(* IEC 61131-3 sources: SortJet_MasterSPS_Aufbau.fbsproj/06_Antriebe/Bosch Rexroth/Rexroth_ctrlX_Drive_Eckelmann_MC_V01_02_02.fb.st^, 26 files *)

(* ---- _Fehlerauswertung.act.st ---- *)
(* METADATA
{
	"v3Meta": {
		"objectGuid": "454009ed-4904-47be-a45e-86d01c03fc0f"
	}
}
*)
ACTION _Fehlerauswertung
/////////////////////////////////////////////////////////////////////////////////////////
/////////////////////////////////////////////////////////////////////////////////////////
// Fehlerauswertung
/////////////////////////////////////////////////////////////////////////////////////////
/////////////////////////////////////////////////////////////////////////////////////////
IF i_ui_Cia402_StatusWord.3 // Fehler am Umrichter aktiv
THEN
  Diagnose := DiagnoseAuswertung( wFehlernummer := udiErrorFromECat );
ELSE
  Diagnose := DiagnoseAuswertung( wFehlernummer := 0 );
END_IF

IF NOT i_ui_Cia402_StatusWord.3 AND NOT blInternerFehler AND blFehlerAktiv AND NOT blFreigabeEntziehenAktiv THEN
  Antriebsfehler.wlBausteinFehlerNr := cMotionFehler;
  blInternerFehler := TRUE;
END_IF

tonlFehlermeldungAusgeben(IN := ( blFehlerAktiv AND Diagnose.bError ) OR blInternerFehler , pt := T#1S);

rtl_Fehlermeldung(CLK := tonlFehlermeldungAusgeben.Q );

bpFehler := blFehlerAktiv AND ( Diagnose.bError (* OR Diagnose.bWarning *) OR blInternerFehler );

IF ( blInternerFehler ) THEN
  wlError := awlFehlerinformationen[4] := DWORD_TO_WORD(Antriebsfehler.wlBausteinFehlerNr);
ELSE
  awlFehlerinformationen[4] := DWORD_TO_WORD(Antriebsfehler.wlAntriebsFehler);
END_IF

IF ( rtl_Fehlermeldung.Q ) THEN

  awlFehlerinformationen[0] := stStationsNummern.NummerExtern;
  awlFehlerinformationen[1] := ppAntriebsInformationen.wpSchaltplanseite;
  awlFehlerinformationen[2] := ppAntriebsInformationen.wpSchaltplanReihe;
  awlFehlerinformationen[3] := ppAntriebsInformationen.wpSchaltschrank;

  IF ( blInternerFehler ) THEN
    SpsError( eFehler_Antrieb,
              wlError,
              stStationsNummern.NummerIntern,
              AutomatikkreisBestimmen(stStationsNummern.NummerSPS),
              awlFehlerinformationen );
  ELSE
    IF ( Diagnose.eType = eRexroth_Fehler_Error ) THEN
      SpsError( eFehler_Rexroth_Fehler + Diagnose.eErrorType,
                Diagnose.wFehlerNr,
                stStationsNummern.NummerIntern,
                AutomatikkreisBestimmen(stStationsNummern.NummerSPS),
                awlFehlerinformationen );
    // Wir loggen keine Warnungen
    // ELSIF ( Diagnose.eType = eRexroth_Fehler_Warning ) THEN
    //   SpsWarnung( eFehler_Rexroth_Warnung + Diagnose.eWarningType,
    //               Diagnose.wFehlerNr,
    //               stStationsNummern.NummerIntern,
    //               AutomatikkreisBestimmen(stStationsNummern.NummerSPS),
    //               awlErrorAdditional );
    END_IF
  END_IF

END_IF
END_ACTION

(* ---- _Statusword.act.st ---- *)
(* METADATA
{
	"v3Meta": {
		"objectGuid": "408b9d1a-1641-4edf-bb35-4e7a7361d31c"
	}
}
*)
ACTION _Statusword
/////////////////////////////////////////////////////////////////////////////////////////
/////////////////////////////////////////////////////////////////////////////////////////
// Aktuellen Status vom Antrieb auslesen
/////////////////////////////////////////////////////////////////////////////////////////
/////////////////////////////////////////////////////////////////////////////////////////
Status();

/////////////////////////////////////////////////////////////////////////////////////////
/////////////////////////////////////////////////////////////////////////////////////////
// Ist-Position auslesen
/////////////////////////////////////////////////////////////////////////////////////////
/////////////////////////////////////////////////////////////////////////////////////////
Istposition();

/////////////////////////////////////////////////////////////////////////////////////////
/////////////////////////////////////////////////////////////////////////////////////////
// Ist-Geschwindigkeit auslesen
/////////////////////////////////////////////////////////////////////////////////////////
/////////////////////////////////////////////////////////////////////////////////////////
IstGeschwindigkeit();

/////////////////////////////////////////////////////////////////////////////////////////
/////////////////////////////////////////////////////////////////////////////////////////
// Hardware Endschalter auslesen
/////////////////////////////////////////////////////////////////////////////////////////
/////////////////////////////////////////////////////////////////////////////////////////
// Rueckmeldung auch bei Quelle SPS aus dem Signal-Statuswort (im Umrichter parametriert)
IF ppAntriebsInformationen.stOptionen.eEndschalterQuelle <> Endschalterquelle_EN.KEINE THEN
  bpMaxSchalterBelegt := i_ui_Signal_StatusWord.1;
  bpMinSchalterBelegt := i_ui_Signal_StatusWord.0;
ELSE
  bpMinSchalterBelegt := FALSE;
  bpMaxSchalterBelegt := FALSE;
END_IF

/////////////////////////////////////////////////////////////////////////////////////////
/////////////////////////////////////////////////////////////////////////////////////////
// Erkennung ob und in welche Richtung der Antrieb verfährt
/////////////////////////////////////////////////////////////////////////////////////////
/////////////////////////////////////////////////////////////////////////////////////////
FahrrichtungErkennung();

/////////////////////////////////////////////////////////////////////////////////////////
/////////////////////////////////////////////////////////////////////////////////////////
// Status-Bits aus Antrieb / Motion holen
/////////////////////////////////////////////////////////////////////////////////////////
/////////////////////////////////////////////////////////////////////////////////////////
IF l_mc_ReadStatus.ErrorStop THEN
  l_mc_ReadAxisError( Axis := ppAntriebsInformationen.wAchsID , Enable := TRUE );
  blReadAxisErrorAktiv := TRUE;
ELSIF blReadAxisErrorAktiv THEN
  l_mc_ReadAxisError( Axis := ppAntriebsInformationen.wAchsID , Enable := FALSE );
  blReadAxisErrorAktiv := FALSE;
END_IF

blFehlerAktiv   := (  i_ui_Cia402_StatusWord.3 // Achsfehler
                     OR ( l_mc_ReadStatus.ErrorStop // MC Fehler
                          AND l_mc_ReadAxisError.Valid
                          AND NOT blFreigabeEntziehenAktiv ) // Aktiver Fehler aus MC_ReadAxisError
                     OR blInternerFehler ); // Fehler im Antriebsbaustein

bpIstReferenziert  := i_ui_Signal_StatusWord.3;
bpAchseSychron     := l_mc_GearIn.InGear (* AND l_mc_ReadStatus.SynchronizedMotion *);
bpBremseGeloest    := i_ui_Signal_StatusWord.15;

blSensoren[eSensoren.Sensor_1] := udipEingaengeUmrichter.cXG31_1_I_1;
blSensoren[eSensoren.Sensor_2] := udipEingaengeUmrichter.cXG31_2_I_2;
blSensoren[eSensoren.Sensor_3] := udipEingaengeUmrichter.cXG31_6_I_4;
blSensoren[eSensoren.Sensor_4] := udipEingaengeUmrichter.cXG31_7_I_5;
blSensoren[eSensoren.Sensor_5] := udipEingaengeUmrichter.cXG37_4_I_6;

// Sensorik vom Slave-gekoppelten Antrieb übernehmen - ggf kann man
IF IsBetweenWORD(wpSlaveNr, 0, 64) AND ( wpSlaveNr <> ppAntriebsInformationen.wAchsID ) THEN
  blSensoren[eSensoren.Sensor_6] := pgAntriebe[wpSlaveNr].udipEingaengeUmrichter.cXG31_1_I_1; // Slave Einlauf
  blSensoren[eSensoren.Sensor_7] := pgAntriebe[wpSlaveNr].udipEingaengeUmrichter.cXG31_2_I_2; // Slave Auslauf
  blSensoren[eSensoren.Sensor_8] := pgAntriebe[wpSlaveNr].udipEingaengeUmrichter.cXG31_6_I_4; // Slave Einlauf Vorab
  blSensoren[eSensoren.Sensor_9] := pgAntriebe[wpSlaveNr].udipEingaengeUmrichter.cXG31_7_I_5; // Slave Auslauf Vorab
ELSE
  blSensoren[eSensoren.Sensor_6] := FALSE;
  blSensoren[eSensoren.Sensor_7] := FALSE;
  blSensoren[eSensoren.Sensor_8] := FALSE;
  blSensoren[eSensoren.Sensor_9] := FALSE;
END_IF

bpMotionAktiv := ( NOT l_mc_ReadStatus.StandStill ) (* OR l_mc_ReadStatus.Disabled *);

bpAntrieblaeuft            := ( eBewegungsrichtung <> TE_Move_Direction.MD_STANDSTILL_E );
bpBewegungsrichtungPositiv := ( eBewegungsrichtung = TE_Move_Direction.MD_POSITIV_E );
bpBewegungsrichtungNegativ := ( eBewegungsrichtung = TE_Move_Direction.MD_NEGATIV_E );

bpKonstantfahrtAktiv       := l_mc_ReadStatus.ConstantVelocity;
bpBeschleunigungAktiv      := l_mc_ReadStatus.Accelerating;
bpVerzoegerungAktiv        := l_mc_ReadStatus.Decelerating;

bpReglerBereit      := ( PowerSupplyStatus.15 AND PowerSupplyStatus.14 AND PowerSupplyStatus.6 AND PowerSupplyStatus.4 )
                       OR ( i_ui_Cia402_StatusWord.0 AND i_ui_Cia402_StatusWord.1 AND i_ui_Cia402_StatusWord.2 );

// Min- und Max-Position bestimmen
rlSoftwareLimitMin := TO_REAL(l_ts_MKAxisConfig.lrSoftwareLimitNegative);
rlSoftwareLimitMax := TO_REAL(l_ts_MKAxisConfig.lrSoftwareLimitPositive);
rpMinPosition := rlSoftwareLimitMin;
rpMaxPosition := rlSoftwareLimitMax;

// Externe Software-Endschalter koennen die MK-Grenzen nur weiter eingrenzen
// 0 bedeutet: kein zusaetzlicher externer Endschalter aktiv

// Min nur enger setzen, nie erweitern
IF rpMinSwEsEingrenzung <> 0 THEN
  IF ( rlSoftwareLimitMin = 0 ) OR ( rpMinSwEsEingrenzung >= rlSoftwareLimitMin ) THEN
    rpMinPosition := rpMinSwEsEingrenzung;
  END_IF
END_IF

// Max nur enger setzen, nie erweitern
IF rpMaxSwEsEingrenzung <> 0 THEN
  IF ( rlSoftwareLimitMax = 0 ) OR ( rpMaxSwEsEingrenzung <= rlSoftwareLimitMax ) THEN
    rpMaxPosition := rpMaxSwEsEingrenzung;
  END_IF
END_IF

// Widerspruch im Ergebnis (Min > Max):
// externe Eingrenzung komplett verwerfen und MK-Grenzen beibehalten
IF rpMinPosition > rpMaxPosition THEN
  rpMinPosition := rlSoftwareLimitMin;
  rpMaxPosition := rlSoftwareLimitMax;
END_IF

blSoftwareLimitAktiv := ( rpMinPosition <> 0 ) OR ( rpMaxPosition <> 0 );

bpAntriebFreigegeben := (     l_mc_Power.Enable
                          AND l_mc_Power.Status );

rpPositionMesstaster1Positiv := TO_REAL(TO_LREAL(diTouchProbe1Pos) / l_ts_MKAxisConfig.lrIncrementsPerDistance * l_ts_MKAxisConfig.lrDistance);
rpPositionMesstaster1Negativ := TO_REAL(TO_LREAL(diTouchProbe1Neg) / l_ts_MKAxisConfig.lrIncrementsPerDistance * l_ts_MKAxisConfig.lrDistance);
rpPositionMesstaster2Positiv := TO_REAL(TO_LREAL(diTouchProbe2Pos) / l_ts_MKAxisConfig.lrIncrementsPerDistance * l_ts_MKAxisConfig.lrDistance);
rpPositionMesstaster2Negativ := TO_REAL(TO_LREAL(diTouchProbe2Neg) / l_ts_MKAxisConfig.lrIncrementsPerDistance * l_ts_MKAxisConfig.lrDistance);

bpHaupschalter400VEin := ppAntriebsInformationen.stOptionen.bVersorgungUeberXVR OR PowerSupplyStatus.4;

/////////////////////////////////////////////////////////////////////////////////////////
/////////////////////////////////////////////////////////////////////////////////////////
// Eingaenge vom Umrichter auslesen
/////////////////////////////////////////////////////////////////////////////////////////
/////////////////////////////////////////////////////////////////////////////////////////
bpLS_150F02_230V := ppAntriebsInformationen.stOptionen.bVersorgungUeberXVR OR udipEingaengeUmrichter.cXG31_3_I_3; // Eingang Leitungsschutzschalter 230V OK

// Ausgangssignale in diesem Normalzyklus uebernehmen, ins Steuerwort schreibt _Steuerwort
wlAusgaengeUmrichter := wpAusgaengeUmrichter;
END_ACTION

(* ---- _Steuerwort.act.st ---- *)
(* METADATA
{
	"v3Meta": {
		"objectGuid": "2cb5236d-2c9d-4e67-a004-d0a59f43b200"
	}
}
*)
ACTION _Steuerwort
// Alle Steuerwort-Bits werden ausschliesslich in dieser Aktion beschrieben.

// Externe Endschalter nur bei Quelle SPS weitergeben, sonst Frei-Pegel (Oeffner: TRUE = frei)
blEndschalterAusSPS := FALSE;
IF __ISVALIDREF(ppAntriebsInformationen) THEN
  blEndschalterAusSPS := ppAntriebsInformationen.stOptionen.eEndschalterQuelle = Endschalterquelle_EN.SPS;
END_IF

SignalSteuerWort.0  := blReferenzLoeschen;
SignalSteuerWort.1  := wlAusgaengeUmrichter.3;
SignalSteuerWort.2  := wlAusgaengeUmrichter.4;
SignalSteuerWort.3  := wlAusgaengeUmrichter.5;
SignalSteuerWort.4  := wlAusgaengeUmrichter.6;
SignalSteuerWort.5  := wlAusgaengeUmrichter.7;
SignalSteuerWort.6  := wlAusgaengeUmrichter.8;
SignalSteuerWort.7  := wlAusgaengeUmrichter.9;
SignalSteuerWort.8  := wlAusgaengeUmrichter.10;
SignalSteuerWort.9  := NOT blEndschalterAusSPS OR bpEndschalterMaxExtern;
SignalSteuerWort.10 := NOT blEndschalterAusSPS OR bpEndschalterMinExtern;
SignalSteuerWort.11 := FALSE;
SignalSteuerWort.12 := FALSE;
SignalSteuerWort.13 := FALSE;
SignalSteuerWort.14 := blReferenzSetzen;
SignalSteuerWort.15 := blBremseLoesen;
END_ACTION

(* ---- A_Changelog.act.st ---- *)
(* METADATA
{
	"v3Meta": {
		"objectGuid": "3ad406ab-889e-4d0d-be2f-76f9c9ecfe4e"
	}
}
*)
{attribute 'excludefrombuild'}
ACTION A_Changelog
(* !!! VERSIONSÄNDERUNGEN WERDEN HIER DETAILLIERT DOKUMENTIERT !!!

- 2025-07-02 - V01_00_00:
  - Entwicklung des Bausteins; Erste Version die Freigegeben wird/wurde

- 2025-10-10 - V01_00_01: Marc Wiegran
  - Änderung des Baustein. Damit die Visualisierung Antriebe_Verfahren weiterhin genutzt werden kann muss in den Schrittketten auf l_mc_power.Enable und nicht auf bpFreigabe geschaut werden.
    l_mc_power.Enable wird aus bpFreigabe und bpFrigabeErzingen, sodass wir nicht mehr in einen Internen Fehler laufen
  - Änderung des Bausteins Damit auch auf die gemeldeten zustände der Hardwarefreigabe geschaut wird wurde in den Schrittketten das l_mc_power.Status durch Regler bereit ersetzt

- 2025-10-15 - V01_00_02: Tobias Brekerbohm
  - Korrektur Vergleich der Software Endschalter - wenn beide 0 dann ansehen als wären keine Aktiv
  - Korrektur bpReglerBereit - Bei Achsen im Zwischenkreis kommen die Bits nicht entsprechend anderer Achsen
    Hier muss auf das CiA Status Word geschaut werden. Zu Prüfen ist, ob das bei den normalen Achsen auch ggf. schon ausreicht
  - Anpassungen / Korrekturen Rotative Achsen

- 2025-10-16 - V01_00_03: Tobias Brekerbohm
  - Korrektur dauernde Neuberechnung der Zielposition bei relativer Positionierung

- 2025-10-17 - V01_00_04: Marc Wiegran
  - Korrektur der Eingangsbits der Langsamfahrnocken auch CoE

- 2025-10-21 - V01_00_05: Marc Wiegran
  - Bei Geschwindigkeitsänderung bei der Messfahrt wird in Step 325 gesprungen um die MC_MOVE_Velocity neu zu starten und nicht wie vorher in 300, da dort erneut die Startbedingungen gepürft werden

- 2025-10-21 - V01_00_06: Marc Wiegran
  - Warteschritt 250 hinzugefgt um sicherzustellen, das die Softwarefreigabe vor Bewegungsstart erteilt wurde noch zu testen ob es die Fehler 6 der MC-Bausteine behebt
  - Schreiben der MC_Home-Fehler-ID in die dafür vorgesehene Variable

- 2025-10-22 - V01_00_07: Marc Wiegran
  - Entfernen des Warteschritt 250, statt dessen wird im Schritt 100 auf l_mc_Power.Status geschaut und Timerüberwacht wird dort ein Fehler ausgeworfen.
      - Enable := Freigabe setzten; Status := Freigabe wurde erfolgreich gesetzt
  - Entfernen der Überprüfung der aktuellen antriebsposition <100 nach der Referenz
      - die Querfahrten haben einen absoluten Referenzoffset von >100, sodass dies andernfalls nicht klappt

- 2025-10-28 - V01_00_08: Tobias Brekerbohm
  - State-Machine achtet nun auf NOT Valid als aller erstes
  - Vergessener Warteschritt 250 aus 1.00.06 der bei der Entfernung in 1.00.07 vergessen wurde zusätzlich entfernt

- 2025-11-11 - V01_00_09: Tobias Brekerbohm
  - Fehlerhaftes ABS setzen von Messergebnissen bei Scheibenmessungen entfernt

- 2025-11-13 - V01_00_10: Tobias Brekerbohm
  - Reset von Ref-Bezug löschen Bit hat gefehlt

- 2025-11-24 - V01_00_11: Tobias Brekerbohm
  - Fehlender Reset von Softwarefreigabe-Timer korigiert
  - An vielen Stellen wurde immernoch auf l_mc_Power.Enable geschaut für den Fehler der Softwarefreigabe statt auf l_mc_Power.Status

- 2026-12-10 - V01_00_12: Tobias Brekerbohm
  - Bei festen Zielpositionen werden keine mm/grad mehr aufaddiert, es werden hart die Grenzwerte aus dem EConSET genommen und nicht mehr schöngerechnet
  - Bei einer Zielpos außerhalb der Grenzen wird nun ein Fehler geworfen, statt die Zielpos stillschweigend zu begrenzen
  - Statt dauernd auf die MK Variablen zu schauen, welche noch konvertiert werden muss, wird nun direkt auf die rpMin- und rpMaxPosition geschaut

- 2026-12-10 - V01_00_13: Tobias Brekerbohm
  - bpAchseSychron schaut nicht länger auf l_mc_ReadStatus.SynchronizedMotion da das Signal aus dem Status gelegentlich geflackert hat

- 2026-12-10 - V01_00_14: Tobias Brekerbohm
  - ReadAxisError wurde nicht aufgerufen
  - Fehlerauswertung bei Fehler aus dem MotionKernel (F 108) bei kein Fehler vom Regler und kein internen Fehler

- 2026-03-12 - V01_00_15: Tobias Brekerbohm
  - Berechnung Ruckzeit bei Langsamfahrt fehlerhaft

- 2026-03-17 - V01_00_16: Tobias Brekerbohm
  - Handplus / Handminus / Restweg-Suchfahrt beachten nun die Software-Endschalter und bremsen vor Erreichen anhand der aktuellen Bremsposition ab
  - Ein Neustart in Richtung eines bereits ueberschrittenen Software-Endschalters wird unterbunden

- 2026-03-19 - V01_00_17: Tobias Brekerbohm
  - Neue Eingaben rpMinSwEsEingrenzung/rpMaxSwEsEingrenzung ergaenzen eine externe Eingrenzung der Software-Endschalter
  - Externe Limits duerfen den MK-Bereich nur enger machen und nicht erweitern
  - Alle Bewegungsarten pruefen neue Zielpositionen und Bremsgrenzen gegen die aktiven Min-/Max-Grenzen

- 2026-03-22 - V01_00_18: Tobias Brekerbohm
  - Antriebssimulation für SPS Simulation (ungetestet)

- 2026-03-24 - V01_00_19: Tobias Brekerbohm
  - XG37-1 und XG37-2 (eigentlich als Eingänge genutzt) optional auch als Ausgänge nutzbar (Benötigt Parameteränderung am Antrieb!!!)

- 2026-03-27 - V01_00_20: Tobias Brekerbohm
  - Neuer Eingang bpFreigabeEntziehenAnhalten fuer kontrollierten Freigabeentzug mit Halt ohne Schrittketten-Reset
  - Bei aktivem Freigabeentzug wird die Achse angehalten, danach die Power entzogen und nach Signalrueckkehr automatisch ohne externen Trigger fortgesetzt
  - Motion-Fehlerauswertung unterdrueckt erwartete ErrorStop-Meldungen waehrend aktivem Freigabeentzug
  - Beim Wiederanlauf nach Freigabeentzug werden laufende Schrittketten auf Execute-Startschritte remappt, damit Bewegungen sicher neu starten
  - Kein ungewollter Schrittketten-Reset bei Signalrueckkehr waehrend aktivem MC_Stop (rtlStop-Kante abgesichert)

- 2026-06-12 - V01_01_00: Tobias Brekerbohm
  - Globaler Override für die Achsgeschwindigkeit - Prozentual zu ändern. Neuer Input rpOverride 0-100
  - Taktzeitoptimierung: Flankenerkennung der Sensoren direkt im Antriebsbaustein ohne zusaetzlichen FB-Aufruf
  - Taktzeitoptimierung: Stillstandsposition nur bei aktiver Software-Endschalter-Bremswegueberwachung berechnen
  - Taktzeitoptimierung: MC_ReadAxisError nur im ErrorStop und einmalig zum Deaktivieren aufrufen
  - S277 Bit 12 wird geprüft, mit Fehlermeldung wenn nicht = 1
  - Bei aktivierter Langsamfahrtnocke wird nicht auf Langsame Geschwindigkeit gestellt, wenn die Achse beim belegen der Nocke/Laser gerade am Verzögern ist.
     Würden wir während der Verzögerung die Geschwindigkeit reduzieren, würde der Verfahrbefehl abgebrochen und neu geschrieben werden in den MotionKernel.
     Dabei verlieren wir Zeit und die Achse würde ihre Zielposition überfahren.
  - Restweg positionierung kann nun auch auf Achsen Restweg fahren, die per wpSlave angegeben werden. Z. b. Greifer auf Riemen-Sensorik (Sensor 6-9)
  - Gravierender Fehler bei der Langsamfahrt behoben: Shuttle überfährt seine Position massiv bei aktiver Langsamfahrt weil die Ruckzeit umgerechnet wurde und dadurch
    die Zielposition nicht mehr erreicht werden kann und somit überschwingt
  - Fehler behoben, dass blInternerFehler erst nach einem 2. Reset zurückgesetzt wurde. MotionFehler brauchten dadurch immer 2 Resets

- 2026-07-07 - V01_01_01: Tobias Brekerbohm
  - Fehler bei Zuweisung von Beschleunigung und Verzögerung behoben.

- 2026-08-04 - V01_01_02: Tobias Brekerbohm
  - Restwegmessung während der Absolutfahrt ermöglicht und Messung mehrerer aufeinanderfolgender Scheiben korrigiert.
  - Messergebnis der Restwegmessung wird immer positiv ausgegeben.

- 2026-08-05 - V01_01_03: Marc Wiegran und Tobias Brekerbohm
  - Korrektur zuweisung rpMessergbnis - Messergebnis war erst einen Zyklus nach erfolgreicher Messung im Statusword
  - Messergebnis der Längenmessung wird wieder negativ ausgegeben, da der Scheibenmessung_FB darauf ausgelegt ist den so zu erhalten

- 2026-09-25 - V01_01_04: Tobias Brekerbohm
  - Langsamfahrt begrenzt die Geschwindigkeit ueber MC_SetOverride auf 10 % der konfigurierten Maximalgeschwindigkeit.
  - Der externe rpOverride bleibt wirksam; Bewegungsbefehle werden fuer Langsamfahrt nicht mehr neu geschrieben.
  - Bei kurz erkanntem Stillstand bleibt aktive Langsamfahrt erhalten, solange eine Langsamfahrtnocke belegt ist.
  - Langsamfahrt-Bedingung in Nockenerkennung, Aktivierung und Halten aufgeteilt; Verhalten unveraendert.

- 2026-10-14 - V01_01_05: Tobias Brekerbohm:
  - FreigabeEntziehen_Wiederanlauf: MC_Stop wird auch ausgeloest, wenn der Antrieb laut MC-Status nicht im Stillstand ist (bisher nur ueber bpAntrieblaeuft -> bei Anlauf/langsamer Fahrt kein Stop und evtl. Power-Entzug waehrend der Fahrt)
  - FreigabeEntziehen_Wiederanlauf: tonlSoftwareFreigabe/tonlHardwareFreigabe werden waehrend des Halts zurueckgesetzt (Haltezeit zaehlt nicht als Timeout der eingefrorenen Schrittkette)

- 2026-10-17 - V01_02_00: Tobias Brekerbohm, Claude
  - Ruck (Jerk) für lineare und rotative Achsen überarbeitet: Kurze Fahrten nutzen von Anfang an den kleineren Jerk. Lange Fahrten starten mit dem Beschleunigungs-Jerk und wechseln bei erreichter Fahrgeschwindigkeit auf den Brems-Jerk. Der Brems-Jerk kann größer oder kleiner sein.
  - Ob eine Fahrt kurz oder lang ist, wird aus Strecke, Geschwindigkeit, Beschleunigung, Verzögerung und Ruckzeit berechnet. Die Ruckzeitbegrenzung aus EConSet wird berücksichtigt.
  - Der Wechsel auf den Brems-Jerk erfolgt nur einmal pro Fahrt. Parameteränderungen und eine Freigabepause schalten nicht wieder in die Beschleunigungsphase zurück.
  - Stoppen verwendet grundsätzlich den Brems-Jerk. Beim Abbruch während der Beschleunigung wird mindestens der Beschleunigungs-Jerk und der Jerk des laufenden Fahrbefehls verwendet. Dieser bleibt bis zum Ende des Stops erhalten, auch wenn die Schrittkette zurückgesetzt wird.
  - Die Jerk-Auswahl wird gemeinsam für Absolut-, Relativ-, Hand-, Mess-, Restweg- und Synchronfahrten verwendet. Strecken werden passend zum Achstyp in Millimetern oder Grad berechnet.

- 2026-10-19 - V01_02_01: Claude
  - Simulation (bgSPS_SIMULATION): MK-Konfiguration wird jetzt auch im Simulationsmodus geladen (MK_GetAxisConfiguration). Vorher blieb l_ts_MKAxisConfig leer und die Achsen liefen mit den Notfall-Grenzen +-1000.
  - Simulation: rlGeschwindigkeit/rlBeschleunigung/rlVerzoegerung werden jetzt wie in Pruefe_Inputs_Langsamfahrt aus den Eingaengen gebildet und auf die MK-Maximalwerte begrenzt. Vorher waren sie im Simulationsmodus immer 0, die Achsen fuhren daher immer mit den Fallback-Werten (200 / 800).
  - Simulation: rpOverride wirkt jetzt auch auf die simulierte Geschwindigkeit.
  - Simulation: Scheibenmessung (SCHEIBENMESSUNG) und Restwegmessung liefern jetzt ein Messergebnis. Mangels Glasmodell gilt eine virtuelle Scheibenlaenge (globale Variable rgSimScheibenlaenge, Standard 1000 mm):
    Die Messung ist abgeschlossen, wenn die Achse seit Messstart (bzw. seit der ersten Flanke bei Restweg) diese Strecke verfahren hat. Vorzeichen wie im Echtbetrieb angenommen: Scheibenmessung negativ (positiv bei bpDrehrichtungsumkehrMessung), Restweg positiv.
    Die Messfahrt laeuft wie im Echtbetrieb immer in positive Richtung. bpMessungOk/bpMessungFehlerhaft/rpMessErgebnis bleiben bis zum Betriebsartenwechsel gespeichert (vorher nur 1 Zyklus).
  - Simulation: Neuer Eingang rpSimMessErgebnis (nur Simulation): Station gibt das Ergebnis der Scheibenmessung vor. Echtbetrieb-Konvention (aus Scheibenmessung_FB): Ergebnis = Scheibenlaenge - Messstrecke, Glaslaenge = ABS(Messstrecke + Ergebnis).
    Die Messfahrt dauert so lange wie der Betrag des Ergebnisses. Ist der Eingang 0, gilt weiter die virtuelle Scheibenlaenge rgSimScheibenlaenge (Vorzeichen negativ).
  - Simulation: bpBremseLoesen setzt SignalSteuerWort.15 (nur mit bpBremseLoesenFreigabe, sonst Fehler) und meldet bpBremseGeloest nach 300 ms zurueck.
  - Simulation: bpAbsolutSetzen durchlaeuft wie im Echtbetrieb Referenz loeschen -> setzen -> bpAbsolutSetzenDone.
  - Simulation: Langsamfahrnocken (bpAktiviereLangsamfahrtNocke) sind jetzt Low-aktiv (FALSE = belegt) wie im Echtbetrieb, an den Wegenden positioniert; bpLangsamfahrenAktiv begrenzt die Geschwindigkeit auf 10 % der MK-Maximalgeschwindigkeit.
  - Simulation: Abbildung Sensor -> Umrichter-Eingang wie im Echtbetrieb (Sensor_3 = XG31_6, Sensor_4 = XG31_7, Sensor_5 = XG37_4; vorher um eine Stelle verschoben). Sensor_6..9 kommen wie im Echtbetrieb vom Slave-Antrieb (wpSlaveNr).

- 2026-10-31 - V01_02_02: Tobias Brekerbohm, Claude
  Hinweis: Die Nummer V01_01_05 wurde in zwei parallelen Zweigen doppelt vergeben: 2026-10-14 TB (FreigabeEntziehen_Wiederanlauf) und 2026-10-06 Daniel Vogelsang.
  Dieser Stand baut auf V01_02_01 auf und uebernimmt die Punkte aus dem zweiten Zweig (V01_01_05 vom 2026-10-06). Ruck-Profil, StopVerwaltung und Simulation bleiben wie in V01_02_01.
  - Steuerwort-Bits zentral in _Steuerwort zusammengefasst; Referenz- und Bremsenbefehle ueber interne BOOL-Merker. _Steuerwort laeuft auch vor den RETURN-Pfaden (ausser Achse 65).
  - Neue Struktur stOptionen (Antrieb_Optionen_ST) in AntriebsInformationen; ersetzt bpHardwareLimits und bpBremseLoesenFreigabe.
  - Endschalterquelle (eEndschalterQuelle): KEINE, UMRICHTER (Signal-Statuswort Bit 0 = Min, Bit 1 = Max) oder SPS.
  - Quelle SPS: Neue Eingaenge bpEndschalterMinExtern/bpEndschalterMaxExtern auf Signal-Steuerwort Bit 10 (Min) und Bit 9 (Max). Oeffner, TRUE = frei, Default TRUE fuer eine nicht vorhandene Seite.
    Bei anderer Quelle bleiben Bit 9/10 auf TRUE. bpMinSchalterBelegt/bpMaxSchalterBelegt kommen auch bei Quelle SPS aus dem Signal-Statuswort.
    Korrektur zum zweiten Zweig: Dort stehen Min/Max in Deklaration und Changelog vertauscht, gesendet wird Bit 9 = Max, Bit 10 = Min.
  - XVR-Modus (bVersorgungUeberXVR): brueckt bpHaupschalter400VEin und bpLS_150F02_230V, ersetzt die festen OR TRUE aus dem zweiten Zweig.
  - BETRIEBSART_MasterSlave Schritt 1000: bpDone wurde per Vergleich gebildet und war dadurch TRUE, obwohl die Achse nicht synchron war bzw. ein Fehler anstand. Jetzt bpDone := l_mc_GearIn.InGear, in den Fehlerzweigen bpDone := FALSE.
  - Defaults setzt bpDone := FALSE. Vorher blieb ein altes bpDone waehrend Busausfall stehen und ein Reset-Auftrag galt sofort als fertig.
  - tonlMaxZeitStatusUngueltig wird jeden Zyklus vor der State Machine aufgerufen und in Defaults zurueckgesetzt. Vorher wurde er nie zurueckgesetzt und eine spaetere kurze Statusstoerung loeste sofort einen Stop aus.
  - BETRIEBSART_Reset Schritt 250: l_mc_Reset.Error wird bewusst nicht ausgewertet. Der Changelog des zweiten Zweigs nennt diesen Punkt, der Code ist dort aber zu Recht auskommentiert.
  - BETRIEBSART_Reset: Neuer Schritt 260, wartet nach MC_Reset 1 s, bevor bei weiter anstehendem Fehler der Reset per CoE laeuft (aus dem zweiten Zweig).
  - _Statusword und Simulation: Widerspruchspruefung der Software-Endschalter auf das Ergebnis (rpMinPosition > rpMaxPosition) umgestellt. Vorher nur, wenn beide externen Grenzen gesetzt waren.
  - Errorstop (AXIS_ERROR_OR_DISABLED mit l_mc_ReadStatus.Errorstop) bricht die aktive Betriebsart ab (ResetStepsUndMcAktionen, Schritt 0, KEINE_FUNKTION, bpDone := FALSE).
    Vorher blieb z. B. HANDPLUS in Schritt 400/1000 mit MoveVelocity.Execute = TRUE stehen, nach dem Reset fehlte die neue Flanke. Ein reines Disabled (Freigabeentzug) behaelt die Schrittkette weiterhin fuer den Wiederanlauf.
  - PruefeFirmwareReferenzBit (S-0-0277 Bit 11): Ein abgebrochener CoE-Lesezugriff wurde als fertig gewertet und meldete mit udiEncoderProperties = 0 faelschlich Fehler 999.
    Jetzt wird nur ein erfolgreiches Lesen ausgewertet; nach Abbruch neuer Versuch nach cTIME_S277_WIEDERHOLEN (10 s), Status in blS277LesenFehlgeschlagen.
    Die Pruefung startet weiterhin erst bei bestehender MMI-Verbindung (Job.tonlMmiOk).
  - CoeReadObject (eigener FB, betrifft l_fb_CoeLesen und l_fb_CoeS277Lesen): ruht im Grundzustand und liest erst nach einer Execute-Flanke.
    Vorher startete der erste Aufruf mit i_b_Execute := FALSE einen Lesezugriff ohne Parameter (EcID 0), was je Achse beim Hochlauf einen PlcError 8002 erzeugte.
    Bei neuem Execute werden o_b_Aborted und der Timeout-Zaehler zurueckgesetzt.
  - BETRIEBSART_MasterSlave Schritt 200: Bei Reglerbereit geht es direkt weiter zu Schritt 400. Der Schritt 300 (Pruefung bpIstReferenziert, Fehler cKeinReferenzpunktBeiPosAbs) entfaellt, ein Slave kann so auch ohne Referenz auf den Master synchronisieren.

*)
END_ACTION

(* ---- BETRIEBSART_Absolut.act.st ---- *)
(* METADATA
{
	"v3Meta": {
		"objectGuid": "4af98741-4e9d-4c0b-ae92-ac6a6c18f571"
	}
}
*)
ACTION BETRIEBSART_Absolut
// Gemeinsame Auswahl; vorhandener Parameter-Re-Entry uebernimmt den Jerk.
rlRuckzeit := RuckFuerBewegung(bStart := asteplSchritt[ABSOLUT] = STEP_450_E,
                                bMitZiel := TRUE, lrZiel := TO_LREAL(rlZielPosition));

CASE asteplSchritt[ABSOLUT] OF

  STEP_0_E:
    IF NOT bpMotionAktiv THEN // Warten bis die Motion nichts anderes aktiv hat
      asteplSchritt[ABSOLUT] := STEP_100_E;
    END_IF

  STEP_100_E:
    tonlSoftwareFreigabe( IN := NOT l_mc_Power.Status, PT := cTIME_HARDWARE_FREIGABE );
    IF l_mc_Power.Status THEN // Nur weitermachen wenn die Software-Freigabe gesetzt ist
      asteplSchritt[ABSOLUT] := STEP_200_E;
    ELSIF tonlSoftwareFreigabe.Q THEN
      asteplSchritt[ABSOLUT] := STEP_900_E;
      blInternerFehler := TRUE;
      Antriebsfehler.wlBausteinFehlerNr := cKeineSoftwareReglerFreigabeBeiPositionierung;
    END_IF

  STEP_200_E:
    tonlHardwareFreigabe( IN := NOT bpReglerBereit, PT := cTIME_HARDWARE_FREIGABE );
    IF bpReglerBereit THEN // Nur weitermachen wenn der Umrichter bereit ist
      asteplSchritt[ABSOLUT] := STEP_300_E;
    ELSIF tonlHardwareFreigabe.Q THEN
      asteplSchritt[ABSOLUT] := STEP_900_E;
      blInternerFehler := TRUE;
      Antriebsfehler.wlBausteinFehlerNr := cKeineHardwareReglerFreigabeBeiPositionierung;
    END_IF

  STEP_300_E:
    IF bpIstReferenziert THEN // Nur weitermachen wenn der Umrichter in Referenz meldet
      asteplSchritt[ABSOLUT] := STEP_400_E;
    ELSE
      asteplSchritt[ABSOLUT] := STEP_900_E;
      blInternerFehler := TRUE;
      Antriebsfehler.wlBausteinFehlerNr := cKeinReferenzpunktBeiPosAbs;
    END_IF

  STEP_400_E:
    // Zielposition überprüfen
    IF blSoftwareLimitAktiv AND ( rpZielposition < rpMinPosition ) THEN
      blInternerFehler := TRUE;
      Antriebsfehler.wlBausteinFehlerNr := cMotionMinimumSoftwareEndschalterAusgeloest;
      asteplSchritt[ABSOLUT] := STEP_900_E;
    ELSIF blSoftwareLimitAktiv AND ( rpZielposition > rpMaxPosition ) THEN
      blInternerFehler := TRUE;
      Antriebsfehler.wlBausteinFehlerNr := cMotionMaximumSoftwareEndschalterAusgeloest;
      asteplSchritt[ABSOLUT] := STEP_900_E;
    ELSE
      rlZielPosition := rpZielposition;
      asteplSchritt[ABSOLUT] := STEP_450_E;
    END_IF

  STEP_450_E:
    l_mc_MoveAbsolute
      (
        Axis := ppAntriebsInformationen.wAchsID,
        Position := rlZielPosition,
        Velocity := rlGeschwindigkeit * cFAKTOR_GESCHWINDIGKEIT,
        Acceleration := rlBeschleunigung * cFAKTOR_RAMPEN,
        Deceleration := rlVerzoegerung * cFAKTOR_RAMPEN,
        Jerk := rlRuckzeit,
        Direction := MC_Direction.MD_SHORTEST_WAY_E,
        BufferMode := MC_BufferMode.BM_ABORTING_E,
        Execute := TRUE
      );

    asteplSchritt[ABSOLUT] := STEP_500_E;

  STEP_500_E:
    IF ( ( ( rlGeschwindigkeit * cFAKTOR_GESCHWINDIGKEIT ) <> l_mc_MoveAbsolute.Velocity )
         OR ( ( rlBeschleunigung * cFAKTOR_RAMPEN ) <> l_mc_MoveAbsolute.Acceleration )
         OR ( ( rlVerzoegerung * cFAKTOR_RAMPEN ) <> l_mc_MoveAbsolute.Deceleration )
         OR (   rlRuckzeit <> l_mc_MoveAbsolute.Jerk ) )
    THEN
      l_mc_MoveAbsolute( Axis := ppAntriebsInformationen.wAchsID, Execute := FALSE );
      asteplSchritt[ABSOLUT] := STEP_400_E;
    ELSIF l_mc_MoveAbsolute.Done AND NOT bpAntrieblaeuft THEN
      l_mc_MoveAbsolute( Axis := ppAntriebsInformationen.wAchsID, Execute := FALSE );
      asteplSchritt[ABSOLUT] := STEP_1000_E;
    ELSIF l_mc_MoveAbsolute.Error THEN
      wlFehlerVonMotionFunktion := l_mc_MoveAbsolute.ErrorID;
      l_mc_MoveAbsolute( Axis := ppAntriebsInformationen.wAchsID, Execute := FALSE );
      asteplSchritt[ABSOLUT] := STEP_900_E;
    END_IF

    l_mc_MoveAbsolute
      (
        Axis := ppAntriebsInformationen.wAchsID
      );

    // Fehler auswertung
    IF NOT l_mc_Power.Status OR NOT bpReglerBereit THEN
      asteplSchritt[ABSOLUT] := STEP_900_E;
      blInternerFehler := TRUE;
      IF NOT l_mc_Power.Status THEN // Nur weitermachen wenn die Software-Freigabe gesetzt ist
        Antriebsfehler.wlBausteinFehlerNr := cKeineSoftwareReglerFreigabeBeiPositionierung;
      ELSE
        Antriebsfehler.wlBausteinFehlerNr := cKeineHardwareReglerFreigabeBeiPositionierung;
      END_IF
    END_IF

  STEP_900_E:
    l_mc_MoveAbsolute( Axis := ppAntriebsInformationen.wAchsID, Execute := FALSE );
    blAchseStoppen := bpReglerBereit AND NOT l_mc_ReadStatus.Errorstop AND ( bpAntrieblaeuft OR bpAchseSychron );

  STEP_1000_E:
    bpDone := TRUE;

END_CASE
END_ACTION

(* ---- BETRIEBSART_Handminus.act.st ---- *)
(* METADATA
{
	"v3Meta": {
		"objectGuid": "6e9ad026-023d-4c36-963c-571344833198"
	}
}
*)
ACTION BETRIEBSART_Handminus
// Gemeinsame Auswahl; vorhandener Parameter-Re-Entry uebernimmt den Jerk.
rlRuckzeit := RuckFuerBewegung(bStart := asteplSchritt[HANDMINUS] = STEP_300_E,
                                bMitZiel := blSoftwareLimitAktiv, lrZiel := TO_LREAL(rpMinPosition));

CASE asteplSchritt[HANDMINUS] OF

  STEP_0_E:
    IF NOT bpMotionAktiv THEN // Warten bis die Motion nichts anderes aktiv hat
      asteplSchritt[HANDMINUS] := STEP_100_E;
    END_IF

  STEP_100_E:
    tonlSoftwareFreigabe( IN := NOT l_mc_Power.Status, PT := cTIME_HARDWARE_FREIGABE );
    IF l_mc_Power.Status THEN // Nur weitermachen wenn die Software-Freigabe gesetzt ist
      asteplSchritt[HANDMINUS] := STEP_200_E;
    ELSIF tonlSoftwareFreigabe.Q THEN
      asteplSchritt[HANDMINUS] := STEP_900_E;
      blInternerFehler := TRUE;
      Antriebsfehler.wlBausteinFehlerNr := cKeineSoftwareReglerFreigabeBeiPositionierung;
    END_IF

  STEP_200_E:
    tonlHardwareFreigabe( IN := NOT bpReglerBereit, PT := cTIME_HARDWARE_FREIGABE );
    IF bpReglerBereit THEN // Nur weitermachen wenn der Umrichter bereit ist
      asteplSchritt[HANDMINUS] := STEP_300_E;
    ELSIF tonlHardwareFreigabe.Q THEN
      asteplSchritt[HANDMINUS] := STEP_900_E;
      blInternerFehler := TRUE;
      Antriebsfehler.wlBausteinFehlerNr := cKeineHardwareReglerFreigabeBeiPositionierung;
    END_IF

  STEP_300_E:
    IF blSoftwareLimitAktiv AND ( rpIstPosition <= rpMinPosition ) THEN
      l_mc_MoveVelocity( Axis := ppAntriebsInformationen.wAchsID, Execute := FALSE );
      blStopOhneReset := TRUE;
      asteplSchritt[HANDMINUS] := STEP_1000_E;
    ELSE
      l_mc_MoveVelocity
        (
          Axis := ppAntriebsInformationen.wAchsID,
          Velocity := rlGeschwindigkeit * cFAKTOR_GESCHWINDIGKEIT,
          Acceleration := rlBeschleunigung * cFAKTOR_RAMPEN,
          Deceleration := rlVerzoegerung * cFAKTOR_RAMPEN,
          Jerk := rlRuckzeit,
          BufferMode := MC_BufferMode.BM_ABORTING_E,
          Direction := MC_Direction.MD_NEGATIV_E,
          Execute := TRUE
        );
      asteplSchritt[HANDMINUS] := STEP_400_E;
    END_IF

  STEP_400_E:
    IF ( ( ( rlGeschwindigkeit * cFAKTOR_GESCHWINDIGKEIT ) <> l_mc_MoveVelocity.Velocity )
         OR ( ( rlBeschleunigung * cFAKTOR_RAMPEN ) <> l_mc_MoveVelocity.Acceleration )
         OR ( ( rlVerzoegerung * cFAKTOR_RAMPEN ) <> l_mc_MoveVelocity.Deceleration )
         OR (   rlRuckzeit <> l_mc_MoveVelocity.Jerk ) )
    THEN
      l_mc_MoveVelocity( Axis := ppAntriebsInformationen.wAchsID, Execute := FALSE );
      asteplSchritt[HANDMINUS] := STEP_300_E;
    ELSIF l_mc_MoveVelocity.Active AND l_mc_MoveVelocity.InVelocity THEN
      l_mc_MoveVelocity( Axis := ppAntriebsInformationen.wAchsID, Execute := FALSE );
      asteplSchritt[HANDMINUS] := STEP_1000_E;
    ELSIF l_mc_MoveVelocity.Error THEN
      wlFehlerVonMotionFunktion := l_mc_MoveVelocity.ErrorID;
      l_mc_MoveVelocity( Axis := ppAntriebsInformationen.wAchsID, Execute := FALSE );
      asteplSchritt[HANDMINUS] := STEP_900_E;
    END_IF

    l_mc_MoveVelocity
      (
        Axis := ppAntriebsInformationen.wAchsID,
      );

    // Fehler auswertung
    IF NOT l_mc_Power.Status OR NOT bpReglerBereit THEN
      asteplSchritt[HANDMINUS] := STEP_900_E;
      blInternerFehler := TRUE;
      IF NOT l_mc_Power.Status THEN // Nur weitermachen wenn die Software-Freigabe gesetzt ist
        Antriebsfehler.wlBausteinFehlerNr := cKeineSoftwareReglerFreigabeBeiPositionierung;
      ELSE
        Antriebsfehler.wlBausteinFehlerNr := cKeineHardwareReglerFreigabeBeiPositionierung;
      END_IF
    END_IF
    IF l_mc_MoveVelocity.Error THEN
      asteplSchritt[HANDMINUS] := STEP_900_E;
    END_IF

    IF    blSoftwareLimitAktiv
          AND ( rlVerzoegerung > 0 )
          AND ( rpStillstandsPosition <= rpMinPosition )
    THEN
      l_mc_MoveVelocity( Axis := ppAntriebsInformationen.wAchsID, Execute := FALSE );
      blStopOhneReset := TRUE;
      blAchseStoppen := bpReglerBereit AND NOT l_mc_ReadStatus.Errorstop AND ( bpAntrieblaeuft OR bpAchseSychron );
      asteplSchritt[HANDMINUS] := STEP_1000_E;
    END_IF

  STEP_900_E:
    l_mc_MoveVelocity( Axis := ppAntriebsInformationen.wAchsID, Execute := FALSE );
    blAchseStoppen := bpReglerBereit AND NOT l_mc_ReadStatus.Errorstop AND ( bpAntrieblaeuft OR bpAchseSychron );

  STEP_1000_E:
    // Fehler auswertung
    IF NOT l_mc_Power.Status OR NOT bpReglerBereit THEN
      asteplSchritt[HANDMINUS] := STEP_900_E;
      blInternerFehler := TRUE;
      IF NOT l_mc_Power.Status THEN // Nur weitermachen wenn die Software-Freigabe gesetzt ist
        Antriebsfehler.wlBausteinFehlerNr := cKeineSoftwareReglerFreigabeBeiPositionierung;
      ELSE
        Antriebsfehler.wlBausteinFehlerNr := cKeineHardwareReglerFreigabeBeiPositionierung;
      END_IF
    END_IF
    IF l_mc_MoveVelocity.Error THEN
      asteplSchritt[HANDMINUS] := STEP_900_E;
    END_IF

    // Parameter geändert ?
    IF ( ( ( rlGeschwindigkeit * cFAKTOR_GESCHWINDIGKEIT ) <> l_mc_MoveVelocity.Velocity )
         OR ( ( rlBeschleunigung * cFAKTOR_RAMPEN ) <> l_mc_MoveVelocity.Acceleration )
         OR ( ( rlVerzoegerung * cFAKTOR_RAMPEN ) <> l_mc_MoveVelocity.Deceleration )
         OR (   rlRuckzeit <> l_mc_MoveVelocity.Jerk ) )
    THEN
      l_mc_MoveVelocity( Axis := ppAntriebsInformationen.wAchsID, Execute := FALSE );
      asteplSchritt[HANDMINUS] := STEP_300_E;
    END_IF

    IF    blSoftwareLimitAktiv
          AND ( rlVerzoegerung > 0 )
          AND ( rpStillstandsPosition <= rpMinPosition )
    THEN
      l_mc_MoveVelocity(Axis := ppAntriebsInformationen.wAchsID, Execute := FALSE);
      blStopOhneReset := TRUE;
      blAchseStoppen := bpReglerBereit AND NOT l_mc_ReadStatus.Errorstop AND ( bpAntrieblaeuft OR bpAchseSychron );
    END_IF

END_CASE
END_ACTION

(* ---- BETRIEBSART_Handplus.act.st ---- *)
(* METADATA
{
	"v3Meta": {
		"objectGuid": "5e7f3be3-98a2-4beb-b625-b580500a4088"
	}
}
*)
ACTION BETRIEBSART_Handplus
// Gemeinsame Auswahl; vorhandener Parameter-Re-Entry uebernimmt den Jerk.
rlRuckzeit := RuckFuerBewegung(bStart := asteplSchritt[HANDPLUS] = STEP_300_E,
                                bMitZiel := blSoftwareLimitAktiv, lrZiel := TO_LREAL(rpMaxPosition));

CASE asteplSchritt[HANDPLUS] OF

  STEP_0_E:
    IF NOT bpMotionAktiv THEN // Warten bis die Motion nichts anderes aktiv hat
      asteplSchritt[HANDPLUS] := STEP_100_E;
    END_IF

  STEP_100_E:
    tonlSoftwareFreigabe( IN := NOT l_mc_Power.Status, PT := cTIME_HARDWARE_FREIGABE );
    IF l_mc_Power.Status THEN // Nur weitermachen wenn die Software-Freigabe gesetzt ist
      asteplSchritt[HANDPLUS] := STEP_200_E;
    ELSIF tonlSoftwareFreigabe.Q THEN
      asteplSchritt[HANDPLUS] := STEP_900_E;
      blInternerFehler := TRUE;
      Antriebsfehler.wlBausteinFehlerNr := cKeineSoftwareReglerFreigabeBeiPositionierung;
    END_IF

  STEP_200_E:
    tonlHardwareFreigabe( IN := NOT bpReglerBereit, PT := cTIME_HARDWARE_FREIGABE );
    IF bpReglerBereit THEN // Nur weitermachen wenn der Umrichter bereit ist
      asteplSchritt[HANDPLUS] := STEP_300_E;
    ELSIF tonlHardwareFreigabe.Q THEN
      asteplSchritt[HANDPLUS] := STEP_900_E;
      blInternerFehler := TRUE;
      Antriebsfehler.wlBausteinFehlerNr := cKeineHardwareReglerFreigabeBeiPositionierung;
    END_IF

  STEP_300_E:
    IF blSoftwareLimitAktiv AND ( rpIstPosition >= rpMaxPosition ) THEN
      l_mc_MoveVelocity( Axis := ppAntriebsInformationen.wAchsID, Execute := FALSE );
      blStopOhneReset := TRUE;
      asteplSchritt[HANDPLUS] := STEP_1000_E;
    ELSE
      l_mc_MoveVelocity
        (
          Axis := ppAntriebsInformationen.wAchsID,
          Velocity := rlGeschwindigkeit * cFAKTOR_GESCHWINDIGKEIT,
          Acceleration := rlBeschleunigung * cFAKTOR_RAMPEN,
          Deceleration := rlVerzoegerung * cFAKTOR_RAMPEN,
          Jerk := rlRuckzeit,
          BufferMode := MC_BufferMode.BM_ABORTING_E,
          Direction := MC_Direction.MD_POSITIV_E,
          Execute := TRUE
        );
      asteplSchritt[HANDPLUS] := STEP_400_E;
    END_IF

  STEP_400_E:
    IF ( ( ( rlGeschwindigkeit * cFAKTOR_GESCHWINDIGKEIT ) <> l_mc_MoveVelocity.Velocity )
         OR ( ( rlBeschleunigung * cFAKTOR_RAMPEN ) <> l_mc_MoveVelocity.Acceleration )
         OR ( ( rlVerzoegerung * cFAKTOR_RAMPEN ) <> l_mc_MoveVelocity.Deceleration )
         OR (   rlRuckzeit <> l_mc_MoveVelocity.Jerk ) )
    THEN
      l_mc_MoveVelocity( Axis := ppAntriebsInformationen.wAchsID, Execute := FALSE );
      asteplSchritt[HANDPLUS] := STEP_300_E;
    ELSIF l_mc_MoveVelocity.Active AND l_mc_MoveVelocity.InVelocity THEN
      l_mc_MoveVelocity( Axis := ppAntriebsInformationen.wAchsID, Execute := FALSE );
      asteplSchritt[HANDPLUS] := STEP_1000_E;
    ELSIF l_mc_MoveVelocity.Error THEN
      wlFehlerVonMotionFunktion := l_mc_MoveVelocity.ErrorID;
      l_mc_MoveVelocity( Axis := ppAntriebsInformationen.wAchsID, Execute := FALSE );
      asteplSchritt[HANDPLUS] := STEP_900_E;
    END_IF

    l_mc_MoveVelocity
      (
        Axis := ppAntriebsInformationen.wAchsID,
      );

    // Fehler auswertung
    IF NOT l_mc_Power.Status OR NOT bpReglerBereit THEN
      asteplSchritt[HANDPLUS] := STEP_900_E;
      blInternerFehler := TRUE;
      IF NOT l_mc_Power.Status THEN // Nur weitermachen wenn die Software-Freigabe gesetzt ist
        Antriebsfehler.wlBausteinFehlerNr := cKeineSoftwareReglerFreigabeBeiPositionierung;
      ELSE
        Antriebsfehler.wlBausteinFehlerNr := cKeineHardwareReglerFreigabeBeiPositionierung;
      END_IF
    END_IF
    IF l_mc_MoveVelocity.Error THEN
      asteplSchritt[HANDPLUS] := STEP_900_E;
    END_IF

    IF     blSoftwareLimitAktiv
           AND ( rlVerzoegerung > 0 )
           AND ( rpStillstandsPosition >= rpMaxPosition )
    THEN
      l_mc_MoveVelocity( Axis := ppAntriebsInformationen.wAchsID, Execute := FALSE );
      blStopOhneReset := TRUE;
      blAchseStoppen := bpReglerBereit AND NOT l_mc_ReadStatus.Errorstop AND ( bpAntrieblaeuft OR bpAchseSychron );
      asteplSchritt[HANDPLUS] := STEP_1000_E;
    END_IF

  STEP_900_E:
    l_mc_MoveVelocity( Axis := ppAntriebsInformationen.wAchsID, Execute := FALSE );
    blAchseStoppen := bpReglerBereit AND NOT l_mc_ReadStatus.Errorstop AND ( bpAntrieblaeuft OR bpAchseSychron );

  STEP_1000_E:
    // Fehler auswertung
    IF NOT l_mc_Power.Status OR NOT bpReglerBereit THEN
      asteplSchritt[HANDPLUS] := STEP_900_E;
      blInternerFehler := TRUE;
      IF NOT l_mc_Power.Status THEN // Nur weitermachen wenn die Software-Freigabe gesetzt ist
        Antriebsfehler.wlBausteinFehlerNr := cKeineSoftwareReglerFreigabeBeiPositionierung;
      ELSE
        Antriebsfehler.wlBausteinFehlerNr := cKeineHardwareReglerFreigabeBeiPositionierung;
      END_IF
    END_IF
    IF l_mc_MoveVelocity.Error THEN
      asteplSchritt[HANDPLUS] := STEP_900_E;
    END_IF

    // Parameter geändert ?
    IF ( ( ( rlGeschwindigkeit * cFAKTOR_GESCHWINDIGKEIT ) <> l_mc_MoveVelocity.Velocity )
         OR ( ( rlBeschleunigung * cFAKTOR_RAMPEN ) <> l_mc_MoveVelocity.Acceleration )
         OR ( ( rlVerzoegerung * cFAKTOR_RAMPEN ) <> l_mc_MoveVelocity.Deceleration )
         OR (   rlRuckzeit <> l_mc_MoveVelocity.Jerk ) )
    THEN
      l_mc_MoveVelocity( Axis := ppAntriebsInformationen.wAchsID, Execute := FALSE );
      asteplSchritt[HANDPLUS] := STEP_300_E;
    END_IF

    IF     blSoftwareLimitAktiv
           AND ( rlVerzoegerung > 0 )
           AND ( rpStillstandsPosition >= rpMaxPosition )
    THEN
      l_mc_MoveVelocity(Axis := ppAntriebsInformationen.wAchsID, Execute := FALSE);
      blStopOhneReset := TRUE;
      blAchseStoppen := bpReglerBereit AND NOT l_mc_ReadStatus.Errorstop AND ( bpAntrieblaeuft OR bpAchseSychron );
    END_IF

END_CASE
END_ACTION

(* ---- BETRIEBSART_MasterSlave.act.st ---- *)
(* METADATA
{
	"v3Meta": {
		"objectGuid": "6d2aa95c-c8c9-48d0-a651-a62b0cc396bc"
	}
}
*)
ACTION BETRIEBSART_MasterSlave
// Gemeinsame Auswahl; vorhandener Parameter-Re-Entry uebernimmt den Jerk.
rlRuckzeit := RuckFuerBewegung(bStart := asteplSchritt[wlSchrittkette] = STEP_400_E,
                                bMitZiel := FALSE, lrZiel := 0);

CASE asteplSchritt[wlSchrittkette] OF

  STEP_0_E:
    IF NOT bpMotionAktiv THEN // Warten bis die Motion nichts anderes aktiv hat
      asteplSchritt[wlSchrittkette] := STEP_100_E;
    END_IF

  STEP_100_E:
    tonlSoftwareFreigabe( IN := NOT l_mc_Power.Status, PT := cTIME_HARDWARE_FREIGABE );
    IF l_mc_Power.Status THEN // Nur weitermachen wenn die Software-Freigabe gesetzt ist
      asteplSchritt[wlSchrittkette] := STEP_200_E;
    ELSIF tonlSoftwareFreigabe.Q THEN
      asteplSchritt[wlSchrittkette] := STEP_900_E;
      blInternerFehler := TRUE;
      Antriebsfehler.wlBausteinFehlerNr := cKeineSoftwareReglerFreigabeBeiPositionierung;
    END_IF

  STEP_200_E:
    tonlHardwareFreigabe( IN := NOT bpReglerBereit, PT := cTIME_HARDWARE_FREIGABE );
    IF bpReglerBereit THEN // Nur weitermachen wenn der Umrichter bereit ist
      asteplSchritt[wlSchrittkette] := STEP_400_E;
    ELSIF tonlHardwareFreigabe.Q THEN
      asteplSchritt[wlSchrittkette] := STEP_900_E;
      blInternerFehler := TRUE;
      Antriebsfehler.wlBausteinFehlerNr := cKeineHardwareReglerFreigabeBeiPositionierung;
    END_IF

  STEP_400_E:
    IF ( NOT IsBetweenWORD(wpMaster, 0, 64) ) OR ( wpMaster = ppAntriebsInformationen.wAchsID ) THEN
      blInternerFehler := TRUE;
      Antriebsfehler.wlBausteinFehlerNr := cBetriebsartNichtUnterstuetzt;
      asteplSchritt[wlSchrittkette] := STEP_900_E;
    ELSE
      l_mc_GearIn
        (
          Slave := ppAntriebsInformationen.wAchsID,
          Master := wpMaster,
          Acceleration := rlBeschleunigung * cFAKTOR_RAMPEN,
          Deceleration := rlVerzoegerung * cFAKTOR_RAMPEN,
          Jerk := rlRuckzeit,
          RatioNumerator := 1,
          RatioDenominator := SEL( ( wlAktiveBetriebsart = INVERTIERTER_SYNC_AUF_MASTER ), 1, -1), // SEL: WENN  ( wlAktiveBetriebsart = INVERTIERTER_SYNC_AUF_MASTER ) = FALSE dann 1 ansonsten -1
          BufferMode := MC_BufferMode.BM_ABORTING_E,
          Execute := TRUE
        );

      asteplSchritt[wlSchrittkette] := STEP_1000_E;
    END_IF

  STEP_900_E:
    l_mc_GearIn( Slave := ppAntriebsInformationen.wAchsID, Master := wpMaster, Execute := FALSE );
    blAchseStoppen := bpReglerBereit AND NOT l_mc_ReadStatus.Errorstop AND ( bpAntrieblaeuft OR bpAchseSychron );

  STEP_1000_E:
    IF ( ( ( rlBeschleunigung * cFAKTOR_RAMPEN ) <> l_mc_GearIn.Acceleration )
         OR ( ( rlVerzoegerung * cFAKTOR_RAMPEN ) <> l_mc_GearIn.Deceleration )
         OR (   rlRuckzeit <> l_mc_GearIn.Jerk ) )
    THEN
      l_mc_GearIn( Slave := ppAntriebsInformationen.wAchsID, Master := wpMaster, Execute := FALSE );
      asteplSchritt[wlSchrittkette] := STEP_400_E;
    END_IF

    l_mc_GearIn
      (
        Slave := ppAntriebsInformationen.wAchsID,
        Master := wpMaster,
      );
    // Done direkt aus dem aktuellen InGear bilden (bpAchseSychron ist der Wert aus dem Vorzyklus)
    bpDone := l_mc_GearIn.InGear;

    // Fehler auswertung
    IF NOT l_mc_Power.Status OR NOT bpReglerBereit THEN
      bpDone := FALSE;
      asteplSchritt[wlSchrittkette] := STEP_900_E;
      blInternerFehler := TRUE;
      IF NOT l_mc_Power.Status THEN // Nur weitermachen wenn die Software-Freigabe gesetzt ist
        Antriebsfehler.wlBausteinFehlerNr := cKeineSoftwareReglerFreigabeBeiPositionierung;
      ELSE
        Antriebsfehler.wlBausteinFehlerNr := cKeineHardwareReglerFreigabeBeiPositionierung;
      END_IF
    END_IF
    IF l_mc_GearIn.Error THEN
      bpDone := FALSE;
      wlFehlerVonMotionFunktion := l_mc_GearIn.ErrorID;
      l_mc_GearIn( Slave := ppAntriebsInformationen.wAchsID, Master := wpMaster, Execute := FALSE );
      asteplSchritt[wlSchrittkette] := STEP_900_E;
    END_IF

END_CASE
END_ACTION

(* ---- BETRIEBSART_Messung.act.st ---- *)
(* METADATA
{
	"v3Meta": {
		"objectGuid": "748a293d-7cb7-4722-9684-4a3f052fb050"
	}
}
*)
ACTION BETRIEBSART_Messung
// Gemeinsame Auswahl; vorhandener Parameter-Re-Entry uebernimmt den Jerk.
rlRuckzeit := RuckFuerBewegung(bStart := asteplSchritt[SCHEIBENMESSUNG] = STEP_325_E,
                                bMitZiel := FALSE, lrZiel := 0);

CASE asteplSchritt[SCHEIBENMESSUNG] OF

  STEP_0_E:
    IF NOT bpMotionAktiv THEN // Warten bis die Motion nichts anderes aktiv hat
      lrlMessenPositionSensor1 := lrlMessenPositionSensor2 := 0.0;
      asteplSchritt[SCHEIBENMESSUNG] := STEP_100_E;
    END_IF

  STEP_100_E:
    tonlSoftwareFreigabe( IN := NOT l_mc_Power.Status, PT := cTIME_HARDWARE_FREIGABE );
    IF l_mc_Power.Status THEN // Nur weitermachen wenn die Software-Freigabe gesetzt ist
      asteplSchritt[SCHEIBENMESSUNG] := STEP_200_E;
    ELSIF tonlSoftwareFreigabe.Q THEN
      asteplSchritt[SCHEIBENMESSUNG] := STEP_900_E;
      blInternerFehler := TRUE;
      Antriebsfehler.wlBausteinFehlerNr := cKeineSoftwareReglerFreigabeBeiPositionierung;
    END_IF

  STEP_200_E:
    tonlHardwareFreigabe( IN := NOT bpReglerBereit, PT := cTIME_HARDWARE_FREIGABE );
    IF bpReglerBereit THEN // Nur weitermachen wenn der Umrichter bereit ist
      asteplSchritt[SCHEIBENMESSUNG] := STEP_300_E;
    ELSIF tonlHardwareFreigabe.Q THEN
      asteplSchritt[SCHEIBENMESSUNG] := STEP_900_E;
      blInternerFehler := TRUE;
      Antriebsfehler.wlBausteinFehlerNr := cKeineHardwareReglerFreigabeBeiPositionierung;
    END_IF

  STEP_300_E:
    IF ( blSensoren[eSensorAuswahl_Messung_1] AND NOT blSensoren[eSensorAuswahl_Messung_2] ) OR ( bpDrehrichtungsumkehrMessung AND NOT blSensoren[eSensorAuswahl_Messung_1] AND blSensoren[eSensorAuswahl_Messung_2] ) THEN
      asteplSchritt[SCHEIBENMESSUNG] := STEP_325_E;
    ELSE
      l_mc_MoveVelocity( Axis := ppAntriebsInformationen.wAchsID, Execute := FALSE );
      bpMessungFehlerhaft := TRUE;
      asteplSchritt[SCHEIBENMESSUNG] := STEP_1000_E;
    END_IF

    // Fehler auswertung
    IF NOT l_mc_Power.Enable OR NOT bpReglerBereit THEN
      asteplSchritt[SCHEIBENMESSUNG] := STEP_900_E;
      blInternerFehler := TRUE;
      IF NOT l_mc_Power.Enable THEN // Nur weitermachen wenn die Software-Freigabe gesetzt ist
        Antriebsfehler.wlBausteinFehlerNr := cKeineSoftwareReglerFreigabeBeiPositionierung;
      ELSE
        Antriebsfehler.wlBausteinFehlerNr := cKeineHardwareReglerFreigabeBeiPositionierung;
      END_IF
    END_IF
    IF l_mc_MoveVelocity.Error THEN
      asteplSchritt[SCHEIBENMESSUNG] := STEP_900_E;
    END_IF

  STEP_325_E:
    l_mc_MoveVelocity
      (
        Axis := ppAntriebsInformationen.wAchsID,
        Velocity := rlGeschwindigkeit * cFAKTOR_GESCHWINDIGKEIT,
        Acceleration := rlBeschleunigung * cFAKTOR_RAMPEN,
        Deceleration := rlVerzoegerung * cFAKTOR_RAMPEN,
        Jerk := rlRuckzeit,
        BufferMode := MC_BufferMode.BM_ABORTING_E,
        Direction := MC_Direction.MD_POSITIV_E,
        Execute := TRUE
      );
    asteplSchritt[SCHEIBENMESSUNG] := STEP_350_E;

  STEP_350_E:

    // Änderungen und Fehler erkennen
    IF ( ( ( rlGeschwindigkeit * cFAKTOR_GESCHWINDIGKEIT ) <> l_mc_MoveVelocity.Velocity )
         OR ( ( rlBeschleunigung * cFAKTOR_RAMPEN ) <> l_mc_MoveVelocity.Acceleration )
         OR ( ( rlVerzoegerung * cFAKTOR_RAMPEN ) <> l_mc_MoveVelocity.Deceleration )
         OR (   rlRuckzeit <> l_mc_MoveVelocity.Jerk ) )
    THEN
      l_mc_MoveVelocity( Axis := ppAntriebsInformationen.wAchsID, Execute := FALSE );
      asteplSchritt[SCHEIBENMESSUNG] := STEP_325_E;
    ELSIF l_mc_MoveVelocity.Active AND l_mc_MoveVelocity.InVelocity THEN
      l_mc_MoveVelocity( Axis := ppAntriebsInformationen.wAchsID, Execute := FALSE );
    ELSIF l_mc_MoveVelocity.Error THEN
      wlFehlerVonMotionFunktion := l_mc_MoveVelocity.ErrorID;
      l_mc_MoveVelocity( Axis := ppAntriebsInformationen.wAchsID, Execute := FALSE );
      asteplSchritt[SCHEIBENMESSUNG] := STEP_900_E;
    END_IF

    l_mc_MoveVelocity
      (
        Axis := ppAntriebsInformationen.wAchsID,
      );

    // Sensorik belegt
    IF bFalling[eSensorAuswahl_Messung_1] THEN
      blMesstaster1Gefunden := TRUE;
      lrlMessenPositionSensor1 := l_mc_ReadActualPosition.Position;
    END_IF
    IF bRising[eSensorAuswahl_Messung_2] THEN
      blMesstaster2Gefunden := TRUE;
      lrlMessenPositionSensor2 := l_mc_ReadActualPosition.Position;
    END_IF

    // Messung vollständig abgeschlossen
    IF blMesstaster1Gefunden AND blMesstaster2Gefunden THEN
      IF NOT bpDrehrichtungsumkehrMessung THEN
        lrlMessErgebnis := (lrlMessenPositionSensor1 - lrlMessenPositionSensor2);
        rpMessErgebnis := TO_REAL(lrlMessErgebnis);
      ELSE
        lrlMessErgebnis := (lrlMessenPositionSensor2 - lrlMessenPositionSensor1);
        rpMessErgebnis := TO_REAL(lrlMessErgebnis);
      END_IF
      bpMessungOk := TRUE;
      blStopOhneReset := TRUE;
      asteplSchritt[SCHEIBENMESSUNG] := STEP_1000_E;
    END_IF

    // Fehler auswertung
    IF NOT l_mc_Power.Enable OR NOT bpReglerBereit THEN
      asteplSchritt[SCHEIBENMESSUNG] := STEP_900_E;
      blInternerFehler := TRUE;
      IF NOT l_mc_Power.Enable THEN // Nur weitermachen wenn die Software-Freigabe gesetzt ist
        Antriebsfehler.wlBausteinFehlerNr := cKeineSoftwareReglerFreigabeBeiPositionierung;
      ELSE
        Antriebsfehler.wlBausteinFehlerNr := cKeineHardwareReglerFreigabeBeiPositionierung;
      END_IF
    END_IF
    IF l_mc_MoveVelocity.Error THEN
      asteplSchritt[SCHEIBENMESSUNG] := STEP_900_E;
    END_IF

  STEP_500_E:
    IF NOT bpAntrieblaeuft AND l_mc_ReadStatus.StandStill THEN
      asteplSchritt[SCHEIBENMESSUNG] := STEP_1000_E;
    END_IF

  STEP_900_E:
    l_mc_MoveVelocity( Axis := ppAntriebsInformationen.wAchsID, Execute := FALSE );
    blAchseStoppen := bpReglerBereit AND NOT l_mc_ReadStatus.Errorstop AND ( bpAntrieblaeuft OR bpAchseSychron );

  STEP_1000_E:
    // Fehler auswertung
    IF NOT l_mc_Power.Status OR NOT bpReglerBereit THEN
      asteplSchritt[SCHEIBENMESSUNG] := STEP_900_E;
      blInternerFehler := TRUE;
      IF NOT l_mc_Power.Status THEN // Nur weitermachen wenn die Software-Freigabe gesetzt ist
        Antriebsfehler.wlBausteinFehlerNr := cKeineSoftwareReglerFreigabeBeiPositionierung;
      ELSE
        Antriebsfehler.wlBausteinFehlerNr := cKeineHardwareReglerFreigabeBeiPositionierung;
      END_IF
    END_IF
    IF l_mc_MoveVelocity.Error THEN
      asteplSchritt[SCHEIBENMESSUNG] := STEP_900_E;
    END_IF

    bpDone := TRUE;

END_CASE
END_ACTION

(* ---- BETRIEBSART_Referenz.act.st ---- *)
(* METADATA
{
	"v3Meta": {
		"objectGuid": "88c040f8-409a-4941-b3a2-808eaede908e"
	}
}
*)
ACTION BETRIEBSART_Referenz
CASE asteplSchritt[REFERENZ] OF

  STEP_0_E:
    IF NOT bpMotionAktiv THEN // Warten bis die Motion nichts anderes aktiv hat
      asteplSchritt[REFERENZ] := STEP_100_E;
    END_IF

  STEP_100_E:

    tonlSoftwareFreigabe( IN := NOT l_mc_Power.Status, PT := cTIME_HARDWARE_FREIGABE );
    IF l_mc_Power.Status THEN // Nur weitermachen wenn die Software-Freigabe gesetzt ist
      blReferenzLoeschen := TRUE; // Referenz ablöschen
      IF NOT bpIstReferenziert THEN
        blReferenzLoeschen := FALSE;
        asteplSchritt[REFERENZ] := STEP_200_E;
      END_IF
    ELSIF tonlSoftwareFreigabe.Q THEN
      asteplSchritt[REFERENZ] := STEP_900_E;
      blInternerFehler := TRUE;
      Antriebsfehler.wlBausteinFehlerNr := cKeineSoftwareReglerFreigabeBeiPositionierung;
    END_IF

  STEP_200_E:
    tonlHardwareFreigabe( IN := NOT bpReglerBereit , PT := cTIME_HARDWARE_FREIGABE );
    IF bpReglerBereit THEN // Nur weitermachen wenn der Umrichter bereit ist
      asteplSchritt[REFERENZ] := STEP_300_E;
    ELSIF tonlHardwareFreigabe.Q THEN
      asteplSchritt[REFERENZ] := STEP_900_E;
      blInternerFehler := TRUE;
      Antriebsfehler.wlBausteinFehlerNr := cKeineHardwareReglerFreigabeBeiPositionierung;
    END_IF

  STEP_300_E:
    // Referenzfahrt ausführen
    l_mc_Home
      (
        Axis := ppAntriebsInformationen.wAchsID,
        Position := 0, //Extra Offset adde to the value of VON_NC.MK,
        Execute := TRUE
      );
    IF l_mc_Home.Done AND bpIstReferenziert AND NOT bpAntrieblaeuft THEN
      l_mc_Home
        (
          Axis := ppAntriebsInformationen.wAchsID,
          Execute := FALSE
        );
      asteplSchritt[REFERENZ] := STEP_1000_E;
    END_IF
    IF l_mc_Home.Error THEN
      wlFehlerVonMotionFunktion := l_mc_Home.ErrorID;
      asteplSchritt[REFERENZ] := STEP_900_E;
    END_IF

    // Fehler auswertung
    IF NOT l_mc_Power.Status OR NOT bpReglerBereit THEN
      asteplSchritt[REFERENZ] := STEP_900_E;
      blInternerFehler := TRUE;
      IF NOT l_mc_Power.Status THEN // Nur weitermachen wenn die Software-Freigabe gesetzt ist
        Antriebsfehler.wlBausteinFehlerNr := cKeineSoftwareReglerFreigabeBeiPositionierung;
      ELSE
        Antriebsfehler.wlBausteinFehlerNr := cKeineHardwareReglerFreigabeBeiPositionierung;
      END_IF
    END_IF

  STEP_900_E:
    l_mc_Home( Axis := ppAntriebsInformationen.wAchsID, Execute := FALSE );
    blAchseStoppen := bpReglerBereit AND NOT l_mc_ReadStatus.Errorstop AND ( bpAntrieblaeuft OR bpAchseSychron );

  STEP_1000_E:
    bpDone := bpIstReferenziert;

END_CASE
END_ACTION

(* ---- BETRIEBSART_Relativ.act.st ---- *)
(* METADATA
{
	"v3Meta": {
		"objectGuid": "7d6d986c-3860-4a6a-9626-b52f70d8fccd"
	}
}
*)
ACTION BETRIEBSART_Relativ
// Gemeinsame Auswahl; vorhandener Parameter-Re-Entry uebernimmt den Jerk.
rlRuckzeit := RuckFuerBewegung(bStart := asteplSchritt[RELATIV] = STEP_400_E,
                                bMitZiel := TRUE, lrZiel := TO_LREAL(rlZielPosition));

CASE asteplSchritt[RELATIV] OF

  STEP_0_E:
    IF NOT bpMotionAktiv THEN // Warten bis die Motion nichts anderes aktiv hat
      asteplSchritt[RELATIV] := STEP_100_E;
    END_IF

  STEP_100_E:
    tonlSoftwareFreigabe( IN := NOT l_mc_Power.Status, PT := cTIME_HARDWARE_FREIGABE );
    IF l_mc_Power.Status THEN // Nur weitermachen wenn die Software-Freigabe gesetzt ist
      asteplSchritt[RELATIV] := STEP_200_E;
    ELSIF tonlSoftwareFreigabe.Q THEN
      asteplSchritt[RELATIV] := STEP_900_E;
      blInternerFehler := TRUE;
      Antriebsfehler.wlBausteinFehlerNr := cKeineSoftwareReglerFreigabeBeiPositionierung;
    END_IF

  STEP_200_E:
    tonlHardwareFreigabe( IN := NOT bpReglerBereit, PT := cTIME_HARDWARE_FREIGABE );
    IF bpReglerBereit THEN // Nur weitermachen wenn der Umrichter bereit ist
      asteplSchritt[RELATIV] := STEP_300_E;//300
    ELSIF tonlHardwareFreigabe.Q THEN
      asteplSchritt[RELATIV] := STEP_900_E;
      blInternerFehler := TRUE;
      Antriebsfehler.wlBausteinFehlerNr := cKeineHardwareReglerFreigabeBeiPositionierung;
    END_IF

  STEP_300_E:
    IF bpIstReferenziert THEN // Nur weitermachen wenn der Umrichter in Referenz meldet
      asteplSchritt[RELATIV] := STEP_350_E;
    ELSE
      asteplSchritt[RELATIV] := STEP_900_E;
      blInternerFehler := TRUE;
      Antriebsfehler.wlBausteinFehlerNr := cKeinReferenzpunktBeiPosAbs;
    END_IF

  STEP_350_E:
    // Für Relativ wird schlicht eine Absolut-Positionierung genutzt
    rlZielposition := rpIstPosition + rpZielposition;

    // Zielposition kleiner/größer Min/max Pos
    IF blSoftwareLimitAktiv AND ( rlZielPosition < rpMinPosition ) THEN
      blInternerFehler := TRUE;
      Antriebsfehler.wlBausteinFehlerNr := cMotionMinimumSoftwareEndschalterAusgeloest;
      asteplSchritt[RELATIV] := STEP_900_E;
    ELSIF blSoftwareLimitAktiv AND ( rlZielPosition > rpMaxPosition ) THEN
      blInternerFehler := TRUE;
      Antriebsfehler.wlBausteinFehlerNr := cMotionMaximumSoftwareEndschalterAusgeloest;
      asteplSchritt[RELATIV] := STEP_900_E;
    ELSE
      asteplSchritt[RELATIV] := STEP_400_E;
    END_IF

  STEP_400_E:

    l_mc_MoveAbsolute
      (
        Axis := ppAntriebsInformationen.wAchsID,
        Position := rlZielposition,
        Velocity := rlGeschwindigkeit * cFAKTOR_GESCHWINDIGKEIT,
        Acceleration := rlBeschleunigung * cFAKTOR_RAMPEN,
        Deceleration := rlVerzoegerung * cFAKTOR_RAMPEN,
        Jerk := rlRuckzeit,
        Direction := MC_Direction.MD_SHORTEST_WAY_E,
        BufferMode := MC_BufferMode.BM_ABORTING_E,
        Execute := TRUE
      );

    asteplSchritt[RELATIV] := STEP_500_E;

  STEP_500_E:
    IF ( ( ( rlGeschwindigkeit * cFAKTOR_GESCHWINDIGKEIT ) <> l_mc_MoveAbsolute.Velocity )
         OR ( ( rlBeschleunigung * cFAKTOR_RAMPEN ) <> l_mc_MoveAbsolute.Acceleration )
         OR ( ( rlVerzoegerung * cFAKTOR_RAMPEN ) <> l_mc_MoveAbsolute.Deceleration )
         OR (   rlRuckzeit <> l_mc_MoveAbsolute.Jerk ) )
    THEN
      l_mc_MoveAbsolute( Axis := ppAntriebsInformationen.wAchsID, Execute := FALSE );
      asteplSchritt[RELATIV] := STEP_400_E;
    ELSIF l_mc_MoveAbsolute.Done THEN
      l_mc_MoveAbsolute( Axis := ppAntriebsInformationen.wAchsID, Execute := FALSE );
      asteplSchritt[RELATIV] := STEP_1000_E;
    ELSIF l_mc_MoveAbsolute.Error THEN
      wlFehlerVonMotionFunktion := l_mc_MoveAbsolute.ErrorID;
      l_mc_MoveAbsolute( Axis := ppAntriebsInformationen.wAchsID, Execute := FALSE );
      asteplSchritt[RELATIV] := STEP_900_E;
    END_IF

    l_mc_MoveAbsolute
      (
        Axis := ppAntriebsInformationen.wAchsID
      );

    // Fehler auswertung
    IF NOT l_mc_Power.Status OR NOT bpReglerBereit THEN
      asteplSchritt[RELATIV] := STEP_900_E;
      blInternerFehler := TRUE;
      IF NOT l_mc_Power.Status THEN // Nur weitermachen wenn die Software-Freigabe gesetzt ist
        Antriebsfehler.wlBausteinFehlerNr := cKeineSoftwareReglerFreigabeBeiPositionierung;
      ELSE
        Antriebsfehler.wlBausteinFehlerNr := cKeineHardwareReglerFreigabeBeiPositionierung;
      END_IF
    END_IF

  STEP_900_E:
    l_mc_MoveAbsolute( Axis := ppAntriebsInformationen.wAchsID, Execute := FALSE );
    blAchseStoppen := bpReglerBereit AND NOT l_mc_ReadStatus.Errorstop AND ( bpAntrieblaeuft OR bpAchseSychron );

  STEP_1000_E:
    bpDone := TRUE;

END_CASE
END_ACTION

(* ---- BETRIEBSART_Reset.act.st ---- *)
(* METADATA
{
	"v3Meta": {
		"objectGuid": "7b92aebb-a3f2-4eb0-b504-974c397a8547"
	}
}
*)
ACTION BETRIEBSART_Reset
CASE asteplSchritt[RESET] OF

  STEP_0_E:
    wlAktiveBetriebsart := RESET;
    ResetStepsUndMcAktionen();
    asteplSchritt[RESET] := STEP_100_E;

  STEP_100_E:
    // Reset nur ausführen WENN Idle und kein Fehler
    // oder Antriebsfehler und dieser Löschbar
    // oder Fehler und kein Fehler vom Antrieb (MC-Error)
    IF ( NOT bpMotionAktiv AND NOT blFehlerAktiv )
       OR ( i_ui_Cia402_StatusWord.3 AND Diagnose.bDeleteable )
       OR ( blFehlerAktiv AND NOT i_ui_Cia402_StatusWord.3 )
       OR ( l_mc_ReadStatus.ErrorStop )
    THEN
      bpFehler                           := FALSE;
      blInternerFehler                   := FALSE;
      wlError                            := 0;
      Diagnose.wFehlerNr                 := 0;
      Antriebsfehler.wlBausteinFehlerNr  := 0;
      tonlFehlermeldungAusgeben(IN := FALSE);
      // l_mc_Power
      // (
      //   Axis   := ppAntriebsInformationen.wAchsID,
      //   Enable := FALSE
      // );
      IF i_ui_Cia402_StatusWord.3 OR l_mc_ReadStatus.ErrorStop THEN
        asteplSchritt[RESET] := STEP_200_E;
      ELSIF NOT blFehlerAktiv THEN
        asteplSchritt[RESET] := STEP_1000_E;
      END_IF
    ELSIF ( i_ui_Cia402_StatusWord.3 AND NOT Diagnose.bDeleteable ) THEN
      bpFehler                           := FALSE;
      blInternerFehler                   := FALSE;
      wlError                            := 0;
      Diagnose.wFehlerNr                 := 0;
      Antriebsfehler.wlBausteinFehlerNr  := 0;
      tonlFehlermeldungAusgeben(IN := FALSE);
      asteplSchritt[RESET] := STEP_1000_E;
    END_IF

  STEP_200_E:
    IF l_mc_ReadStatus.Errorstop THEN
      l_mc_Reset(
                  Axis := ppAntriebsInformationen.wAchsID,
                  Execute := TRUE
                );
      asteplSchritt[RESET] := STEP_250_E;
    ELSE
      IF i_ui_Cia402_StatusWord.3 THEN
        asteplSchritt[RESET] := STEP_275_E;
      ELSE
        blInternerFehler := FALSE;
        Antriebsfehler.wlBausteinFehlerNr := 0;
        asteplSchritt[RESET] := STEP_1000_E;
      END_IF
    END_IF

  STEP_250_E:
    l_mc_Reset(
                Axis := ppAntriebsInformationen.wAchsID
              );
    IF l_mc_Reset.Done THEN
      l_mc_Reset(
                  Axis := ppAntriebsInformationen.wAchsID,
                  Execute := FALSE
                );
      IF i_ui_Cia402_StatusWord.3 THEN
        tonlWarteAufReset( IN := FALSE );
        asteplSchritt[RESET] := STEP_260_E;
      ELSE
        blInternerFehler := FALSE;
        Antriebsfehler.wlBausteinFehlerNr := 0;
        asteplSchritt[RESET] := STEP_1000_E;
      END_IF
    END_IF

  STEP_260_E:
    // Dem Antrieb Zeit geben, den Fehler nach MC_Reset selbst zu loeschen
    tonlWarteAufReset( IN := TRUE, PT := T#1S );
    IF tonlWarteAufReset.Q THEN
      tonlWarteAufReset( IN := FALSE );
      asteplSchritt[RESET] := STEP_275_E;
    END_IF

  //
  // RESET VIA CoE Write
  //
  STEP_275_E:
    l_fb_CoeSchreiben( i_by_EcID := 1000+l_ts_MKAxisConfig.uiDeviceAddress, i_b_Execute := FALSE, i_b_Reset := TRUE );
    IF NOT l_fb_CoeSchreiben.o_b_Busy THEN
      asteplSchritt[RESET] := STEP_300_E;
    END_IF

  STEP_300_E:
    uilSchreibeUeberCoe := 3;
    l_fb_CoeSchreiben
      (
        i_by_EcID      := 1000+l_ts_MKAxisConfig.uiDeviceAddress,
        i_w_ObjectNum  := 16#2B87,
        i_by_SubIndex  := 2,
        i_w_DataTyp    := 6,
        i_p_Var        := ADR(uilSchreibeUeberCoe),
        i_w_BufSize    := SIZEOF(uilSchreibeUeberCoe)
      );
    l_fb_CoeSchreiben( i_b_Execute := TRUE );
    asteplSchritt[RESET] := STEP_325_E;

  STEP_325_E:
    l_fb_CoeSchreiben();
    IF l_fb_CoeSchreiben.o_b_Busy THEN
      asteplSchritt[RESET] := STEP_350_E;
    END_IF

  STEP_350_E:
    l_fb_CoeSchreiben();
    IF NOT l_fb_CoeSchreiben.o_b_Busy THEN
      asteplSchritt[RESET] := STEP_400_E;
    END_IF

  STEP_400_E:
    l_fb_CoeSchreiben( i_by_EcID := 1000+l_ts_MKAxisConfig.uiDeviceAddress, i_b_Execute := FALSE, i_b_Reset := TRUE );
    IF NOT l_fb_CoeSchreiben.o_b_Busy THEN
      asteplSchritt[RESET] := STEP_450_E;
    END_IF

  STEP_450_E:
    uilSchreibeUeberCoe := 0;
    l_fb_CoeSchreiben
      (
        i_by_EcID      := 1000+l_ts_MKAxisConfig.uiDeviceAddress,
        i_w_ObjectNum  := 16#2B87,
        i_by_SubIndex  := 2,
        i_w_DataTyp    := 6,
        i_p_Var        := ADR(uilSchreibeUeberCoe),
        i_w_BufSize    := SIZEOF(uilSchreibeUeberCoe)
      );
    l_fb_CoeSchreiben( i_b_Execute := TRUE );
    asteplSchritt[RESET] := STEP_475_E;

  STEP_475_E:
    l_fb_CoeSchreiben();
    IF l_fb_CoeSchreiben.o_b_Busy THEN
      asteplSchritt[RESET] := STEP_500_E;
    END_IF

  STEP_500_E:
    l_fb_CoeSchreiben();
    IF NOT l_fb_CoeSchreiben.o_b_Busy THEN
      blInternerFehler := FALSE;
      Antriebsfehler.wlBausteinFehlerNr := 0;
      asteplSchritt[RESET] := STEP_1000_E;
    END_IF

  STEP_1000_E:
    wlAktiveBetriebsart := KEINE_FUNKTION;
    bpDone := NOT bpFehler OR NOT Diagnose.bDeleteable;

END_CASE
END_ACTION

(* ---- BETRIEBSART_Restweg_Mit_Messung.act.st ---- *)
(* METADATA
{
	"v3Meta": {
		"objectGuid": "2ee0d1a4-84c9-4083-9399-00f06b07a933"
	}
}
*)
ACTION BETRIEBSART_Restweg_Mit_Messung
// Gemeinsame Auswahl; vorhandener Parameter-Re-Entry uebernimmt den Jerk.
rlRuckzeit := RuckFuerBewegung(bStart := (asteplSchritt[RESTWEG] = STEP_400_E)
                                OR (asteplSchritt[RESTWEG] = STEP_525_E),
                                bMitZiel := asteplSchritt[RESTWEG] >= STEP_500_E,
                                lrZiel := TO_LREAL(rlZielPosition));

CASE asteplSchritt[RESTWEG] OF

  STEP_0_E:
    IF NOT bpMotionAktiv THEN // Warten bis die Motion nichts anderes aktiv hat
      asteplSchritt[RESTWEG] := STEP_100_E;
    END_IF

  STEP_100_E:
    tonlSoftwareFreigabe( IN := NOT l_mc_Power.Status, PT := cTIME_HARDWARE_FREIGABE );
    IF l_mc_Power.Status THEN // Nur weitermachen wenn die Software-Freigabe gesetzt ist
      asteplSchritt[RESTWEG] := STEP_200_E;
    ELSIF tonlSoftwareFreigabe.Q THEN
      asteplSchritt[RESTWEG] := STEP_900_E;
      blInternerFehler := TRUE;
      Antriebsfehler.wlBausteinFehlerNr := cKeineSoftwareReglerFreigabeBeiPositionierung;
    END_IF

  STEP_200_E:
    tonlHardwareFreigabe( IN := NOT bpReglerBereit, PT := cTIME_HARDWARE_FREIGABE );
    IF bpReglerBereit THEN // Nur weitermachen wenn der Umrichter bereit ist
      asteplSchritt[RESTWEG] := STEP_300_E;
    ELSIF tonlHardwareFreigabe.Q THEN
      asteplSchritt[RESTWEG] := STEP_900_E;
      blInternerFehler := TRUE;
      Antriebsfehler.wlBausteinFehlerNr := cKeineHardwareReglerFreigabeBeiPositionierung;
    END_IF

  STEP_300_E:
    IF bpIstReferenziert THEN // Nur weitermachen wenn der Umrichter in Referenz meldet
      asteplSchritt[RESTWEG] := STEP_400_E;
    ELSE
      asteplSchritt[RESTWEG] := STEP_900_E;
      blInternerFehler := TRUE;
      Antriebsfehler.wlBausteinFehlerNr := cKeinReferenzpunktBeiPosAbs;
    END_IF

  STEP_400_E:
    // Drehrichtung für Suchfahrt bestimmen
    IF wpRestwegMode.0 THEN
      l_mc_MoveVelocity.Direction :=  MC_Direction.MD_POSITIV_E;
    ELSE
      l_mc_MoveVelocity.Direction :=  MC_Direction.MD_NEGATIV_E;
    END_IF

    IF wpRestwegMode.0 AND blSoftwareLimitAktiv AND ( rpIstPosition >= rpMaxPosition ) THEN
      blInternerFehler := TRUE;
      Antriebsfehler.wlBausteinFehlerNr := cMotionMaximumSoftwareEndschalterAusgeloest;
      blStopOhneReset := TRUE;
      asteplSchritt[RESTWEG] := STEP_900_E;
    ELSIF ( NOT wpRestwegMode.0 ) AND blSoftwareLimitAktiv AND ( rpIstPosition <= rpMinPosition ) THEN
      blInternerFehler := TRUE;
      Antriebsfehler.wlBausteinFehlerNr := cMotionMinimumSoftwareEndschalterAusgeloest;
      blStopOhneReset := TRUE;
      asteplSchritt[RESTWEG] := STEP_900_E;
    ELSE
      l_mc_MoveVelocity
        (
          Axis := ppAntriebsInformationen.wAchsID,
          Velocity := rlGeschwindigkeit * cFAKTOR_GESCHWINDIGKEIT,
          Acceleration := rlBeschleunigung * cFAKTOR_RAMPEN,
          Deceleration := rlVerzoegerung * cFAKTOR_RAMPEN,
          Jerk := rlRuckzeit,
          BufferMode := MC_BufferMode.BM_ABORTING_E,
          Execute := TRUE
        );
      asteplSchritt[RESTWEG] := STEP_450_E;
    END_IF

    // Sensorik prüfen für Flanken und Messung
    BETRIEBSART_Restweg_X_Flankenerkennung();

  STEP_450_E:
    // Fahrparameter geändert
    IF ( ( ( rlGeschwindigkeit * cFAKTOR_GESCHWINDIGKEIT ) <> l_mc_MoveVelocity.Velocity )
         OR ( ( rlBeschleunigung * cFAKTOR_RAMPEN ) <> l_mc_MoveVelocity.Acceleration )
         OR ( ( rlVerzoegerung * cFAKTOR_RAMPEN ) <> l_mc_MoveVelocity.Deceleration )
         OR (   rlRuckzeit <> l_mc_MoveVelocity.Jerk ) )
    THEN
      l_mc_MoveVelocity( Axis := ppAntriebsInformationen.wAchsID, Execute := FALSE );
      asteplSchritt[RESTWEG] := STEP_400_E;
    ELSIF l_mc_MoveVelocity.Error THEN
      wlFehlerVonMotionFunktion := l_mc_MoveVelocity.ErrorID;
      l_mc_MoveVelocity( Axis := ppAntriebsInformationen.wAchsID, Execute := FALSE );
      asteplSchritt[RESTWEG] := STEP_900_E;
    END_IF

    l_mc_MoveVelocity
      (
        Axis := ppAntriebsInformationen.wAchsID,
      );

    IF ( rlVerzoegerung > 0 ) THEN
      IF    wpRestwegMode.0
            AND blSoftwareLimitAktiv
            AND ( rpStillstandsPosition >= rpMaxPosition )
      THEN
        blInternerFehler := TRUE;
        Antriebsfehler.wlBausteinFehlerNr := cMotionMaximumSoftwareEndschalterAusgeloest;
        l_mc_MoveVelocity( Axis := ppAntriebsInformationen.wAchsID, Execute := FALSE );
        blStopOhneReset := TRUE;
        blAchseStoppen := bpReglerBereit AND NOT l_mc_ReadStatus.Errorstop AND ( bpAntrieblaeuft OR bpAchseSychron );
        asteplSchritt[RESTWEG] := STEP_900_E;
      ELSIF ( NOT wpRestwegMode.0 )
            AND blSoftwareLimitAktiv
            AND ( rpStillstandsPosition <= rpMinPosition )
      THEN
        blInternerFehler := TRUE;
        Antriebsfehler.wlBausteinFehlerNr := cMotionMinimumSoftwareEndschalterAusgeloest;
        l_mc_MoveVelocity( Axis := ppAntriebsInformationen.wAchsID, Execute := FALSE );
        blStopOhneReset := TRUE;
        blAchseStoppen := bpReglerBereit AND NOT l_mc_ReadStatus.Errorstop AND ( bpAntrieblaeuft OR bpAchseSychron );
        asteplSchritt[RESTWEG] := STEP_900_E;
      ELSE
        // Sensorik prüfen für Flanken und Messung
        BETRIEBSART_Restweg_X_Flankenerkennung();
      END_IF
    ELSE
      // Sensorik prüfen für Flanken und Messung
      BETRIEBSART_Restweg_X_Flankenerkennung();
    END_IF

  STEP_500_E:
    bpRestwegMaterialGefunden := TRUE;
    rlZielPosition := TO_REAL(lrlRestwegMesstasterGefunden) + rpZielPosition;

    // Sensorik weiterhin für die Messung auswerten
    BETRIEBSART_Restweg_X_Flankenerkennung();

    // Zielposition kleiner/größer Min/max Pos
    IF blSoftwareLimitAktiv AND ( rlZielPosition < rpMinPosition ) THEN
      blInternerFehler := TRUE;
      Antriebsfehler.wlBausteinFehlerNr := cMotionMinimumSoftwareEndschalterAusgeloest;
      asteplSchritt[RESTWEG] := STEP_900_E;
    ELSIF blSoftwareLimitAktiv AND ( rlZielPosition > rpMaxPosition ) THEN
      blInternerFehler := TRUE;
      Antriebsfehler.wlBausteinFehlerNr := cMotionMaximumSoftwareEndschalterAusgeloest;
      asteplSchritt[RESTWEG] := STEP_900_E;
    ELSE
      asteplSchritt[RESTWEG] := STEP_525_E;
    END_IF

  STEP_525_E:
    l_mc_MoveAbsolute
      (
        Axis := ppAntriebsInformationen.wAchsID,
        Position := rlZielPosition,
        Velocity := rlGeschwindigkeit * cFAKTOR_GESCHWINDIGKEIT,
        Acceleration := rlBeschleunigung * cFAKTOR_RAMPEN,
        Deceleration := rlVerzoegerung * cFAKTOR_RAMPEN,
        Jerk := rlRuckzeit,
        Direction := MC_Direction.MD_SHORTEST_WAY_E,
        BufferMode := MC_BufferMode.BM_ABORTING_E,
        Execute := TRUE
      );

    // Sensorik weiterhin für die Messung auswerten
    BETRIEBSART_Restweg_X_Flankenerkennung();

    asteplSchritt[RESTWEG] := STEP_550_E;

  STEP_550_E:
    IF ( ( ( rlGeschwindigkeit * cFAKTOR_GESCHWINDIGKEIT ) <> l_mc_MoveAbsolute.Velocity )
         OR ( ( rlBeschleunigung * cFAKTOR_RAMPEN ) <> l_mc_MoveAbsolute.Acceleration )
         OR ( ( rlVerzoegerung * cFAKTOR_RAMPEN ) <> l_mc_MoveAbsolute.Deceleration )
         OR (   rlRuckzeit <> l_mc_MoveAbsolute.Jerk ) )
    THEN
      l_mc_MoveAbsolute( Axis := ppAntriebsInformationen.wAchsID, Execute := FALSE );
      asteplSchritt[RESTWEG] := STEP_500_E;
    ELSIF l_mc_MoveAbsolute.Done AND NOT bpAntrieblaeuft THEN
      l_mc_MoveAbsolute( Axis := ppAntriebsInformationen.wAchsID, Execute := FALSE );
      asteplSchritt[RESTWEG] := STEP_1000_E;
    ELSIF l_mc_MoveAbsolute.Error THEN
      wlFehlerVonMotionFunktion := l_mc_MoveAbsolute.ErrorID;
      l_mc_MoveAbsolute( Axis := ppAntriebsInformationen.wAchsID, Execute := FALSE );
      asteplSchritt[RESTWEG] := STEP_900_E;
    END_IF

    l_mc_MoveAbsolute
      (
        Axis := ppAntriebsInformationen.wAchsID
      );

    // Während der gesamten Absolutfahrt die zweite Flanke erfassen
    BETRIEBSART_Restweg_X_Flankenerkennung();

    // Fehler auswertung
    IF NOT l_mc_Power.Status OR NOT bpReglerBereit THEN
      asteplSchritt[RESTWEG] := STEP_900_E;
      blInternerFehler := TRUE;
      IF NOT l_mc_Power.Status THEN // Nur weitermachen wenn die Software-Freigabe gesetzt ist
        Antriebsfehler.wlBausteinFehlerNr := cKeineSoftwareReglerFreigabeBeiPositionierung;
      ELSE
        Antriebsfehler.wlBausteinFehlerNr := cKeineHardwareReglerFreigabeBeiPositionierung;
      END_IF
    END_IF

  STEP_900_E:
    l_mc_MoveVelocity( Axis := ppAntriebsInformationen.wAchsID, Execute := FALSE );
    l_mc_MoveAbsolute( Axis := ppAntriebsInformationen.wAchsID, Execute := FALSE );
    blAchseStoppen := bpReglerBereit AND NOT l_mc_ReadStatus.Errorstop AND ( bpAntrieblaeuft OR bpAchseSychron );

  STEP_1000_E:
    bpDone := TRUE;

END_CASE
END_ACTION

(* ---- BETRIEBSART_Restweg_X_Flankenerkennung.act.st ---- *)
(* METADATA
{
	"v3Meta": {
		"objectGuid": "1c89a038-43c8-45ac-ae17-8c8fe5411e58"
	}
}
*)
ACTION BETRIEBSART_Restweg_X_Flankenerkennung
/////////////////////////////////////////////////////////////////////////////////////////
/////////////////////////////////////////////////////////////////////////////////////////
// RESTWEG - SUCHFAHRT
/////////////////////////////////////////////////////////////////////////////////////////
/////////////////////////////////////////////////////////////////////////////////////////
IF (  asteplSchritt[RESTWEG] < STEP_500_E
     AND asteplSchritt[RESTWEG] > STEP_399_E )
THEN

  IF wpRestwegMode.4 THEN // Steigende Flanke !!!

    IF ( wpRestwegMode.2 AND bRising[eSensoren.Sensor_1] )
       OR ( wpRestwegMode.3 AND bRising[eSensoren.Sensor_2] )
       OR ( wpRestwegMode.5 AND bRising[eSensoren.Sensor_3] )
       OR ( wpRestwegMode.6 AND bRising[eSensoren.Sensor_4] )
       OR ( wpRestwegMode.7 AND bRising[eSensoren.Sensor_5] )
       OR ( wpRestwegMode.8 AND bRising[eSensoren.Sensor_6] )
       OR ( wpRestwegMode.9 AND bRising[eSensoren.Sensor_7] )
       OR ( wpRestwegMode.10 AND bRising[eSensoren.Sensor_8] )
       OR ( wpRestwegMode.11 AND bRising[eSensoren.Sensor_9] )
    THEN
      lrlRestwegMessungMesstasterGefunden := lrlRestwegMesstasterGefunden := l_mc_ReadActualPosition.Position;
      blHelfer_RestwegMesung_Objekt_Gefunden := TRUE;
      l_mc_MoveVelocity( Axis := ppAntriebsInformationen.wAchsID, Execute := FALSE );
      asteplSchritt[RESTWEG] := STEP_500_E;
    END_IF

  ELSE // Fallende Flanke

    IF ( wpRestwegMode.2 AND bFalling[eSensoren.Sensor_1] )
       OR ( wpRestwegMode.3 AND bFalling[eSensoren.Sensor_2] )
       OR ( wpRestwegMode.5 AND bFalling[eSensoren.Sensor_3] )
       OR ( wpRestwegMode.6 AND bFalling[eSensoren.Sensor_4] )
       OR ( wpRestwegMode.7 AND bFalling[eSensoren.Sensor_5] )
       OR ( wpRestwegMode.8 AND bFalling[eSensoren.Sensor_6] )
       OR ( wpRestwegMode.9 AND bFalling[eSensoren.Sensor_7] )
       OR ( wpRestwegMode.10 AND bFalling[eSensoren.Sensor_8] )
       OR ( wpRestwegMode.11 AND bFalling[eSensoren.Sensor_9] )
    THEN
      lrlRestwegMessungMesstasterGefunden := lrlRestwegMesstasterGefunden := l_mc_ReadActualPosition.Position;
      blHelfer_RestwegMesung_Objekt_Gefunden := TRUE;
      l_mc_MoveVelocity( Axis := ppAntriebsInformationen.wAchsID, Execute := FALSE );
      asteplSchritt[RESTWEG] := STEP_500_E;
    END_IF

  END_IF

END_IF

/////////////////////////////////////////////////////////////////////////////////////////
/////////////////////////////////////////////////////////////////////////////////////////
// AUSWERTUNG MESSUNG
/////////////////////////////////////////////////////////////////////////////////////////
/////////////////////////////////////////////////////////////////////////////////////////

IF ( asteplSchritt[RESTWEG] >= STEP_500_E ) THEN

  // (neues) Objekt wurde gefunden
  IF blHelfer_RestwegMesung_Objekt_Gefunden THEN

    // Restweg ursprünglich auf steigende Flanke - jetzt auf fallende Flanke warten
    IF wpRestwegMode.4 THEN // Steigende Flanke !!!

      IF ( wpRestwegMode.2 AND bFalling[eSensoren.Sensor_1] )
         OR ( wpRestwegMode.3 AND bFalling[eSensoren.Sensor_2] )
         OR ( wpRestwegMode.5 AND bFalling[eSensoren.Sensor_3] )
         OR ( wpRestwegMode.6 AND bFalling[eSensoren.Sensor_4] )
         OR ( wpRestwegMode.7 AND bFalling[eSensoren.Sensor_5] )
         OR ( wpRestwegMode.8 AND bFalling[eSensoren.Sensor_6] )
         OR ( wpRestwegMode.9 AND bFalling[eSensoren.Sensor_7] )
         OR ( wpRestwegMode.10 AND bFalling[eSensoren.Sensor_8] )
         OR ( wpRestwegMode.11 AND bFalling[eSensoren.Sensor_9] )
      THEN
        lrlMessErgebnis := ABS(l_mc_ReadActualPosition.Position - lrlRestwegMessungMesstasterGefunden);
        rpMessErgebnis := TO_REAL(lrlMessErgebnis);
        bpMessungOk := TRUE;
        blHelfer_RestwegMesung_Objekt_Gefunden := FALSE;
      END_IF

    // Restweg ursprünglich auf fallende Flanke - jetzt auf steigende Flanke warten
    ELSE // Fallende Flanke

      IF ( wpRestwegMode.2 AND bRising[eSensoren.Sensor_1] )
         OR ( wpRestwegMode.3 AND bRising[eSensoren.Sensor_2] )
         OR ( wpRestwegMode.5 AND bRising[eSensoren.Sensor_3] )
         OR ( wpRestwegMode.6 AND bRising[eSensoren.Sensor_4] )
         OR ( wpRestwegMode.7 AND bRising[eSensoren.Sensor_5] )
         OR ( wpRestwegMode.8 AND bRising[eSensoren.Sensor_6] )
         OR ( wpRestwegMode.9 AND bRising[eSensoren.Sensor_7] )
         OR ( wpRestwegMode.10 AND bRising[eSensoren.Sensor_8] )
         OR ( wpRestwegMode.11 AND bRising[eSensoren.Sensor_9] )
      THEN
        lrlMessErgebnis := ABS(l_mc_ReadActualPosition.Position - lrlRestwegMessungMesstasterGefunden);
        rpMessErgebnis := TO_REAL(lrlMessErgebnis);
        bpMessungOk := TRUE;
        blHelfer_RestwegMesung_Objekt_Gefunden := FALSE;
      END_IF

    END_IF

  // Objekt noch nicht gefunden
  ELSE

    IF wpRestwegMode.4 THEN // Steigende Flanke !!!

      IF ( wpRestwegMode.2 AND bRising[eSensoren.Sensor_1] )
         OR ( wpRestwegMode.3 AND bRising[eSensoren.Sensor_2] )
         OR ( wpRestwegMode.5 AND bRising[eSensoren.Sensor_3] )
         OR ( wpRestwegMode.6 AND bRising[eSensoren.Sensor_4] )
         OR ( wpRestwegMode.7 AND bRising[eSensoren.Sensor_5] )
         OR ( wpRestwegMode.8 AND bRising[eSensoren.Sensor_6] )
         OR ( wpRestwegMode.9 AND bRising[eSensoren.Sensor_7] )
         OR ( wpRestwegMode.10 AND bRising[eSensoren.Sensor_8] )
         OR ( wpRestwegMode.11 AND bRising[eSensoren.Sensor_9] )
      THEN
        lrlMessErgebnis := rpMessErgebnis := 0;
        bpMessungOk := FALSE;
        blHelfer_RestwegMesung_Objekt_Gefunden := TRUE;
        lrlRestwegMessungMesstasterGefunden := l_mc_ReadActualPosition.Position;
      END_IF

    ELSE // Fallende Flanke

      IF ( wpRestwegMode.2 AND bFalling[eSensoren.Sensor_1] )
         OR ( wpRestwegMode.3 AND bFalling[eSensoren.Sensor_2] )
         OR ( wpRestwegMode.5 AND bFalling[eSensoren.Sensor_3] )
         OR ( wpRestwegMode.6 AND bFalling[eSensoren.Sensor_4] )
         OR ( wpRestwegMode.7 AND bFalling[eSensoren.Sensor_5] )
         OR ( wpRestwegMode.8 AND bFalling[eSensoren.Sensor_6] )
         OR ( wpRestwegMode.9 AND bFalling[eSensoren.Sensor_7] )
         OR ( wpRestwegMode.10 AND bFalling[eSensoren.Sensor_8] )
         OR ( wpRestwegMode.11 AND bFalling[eSensoren.Sensor_9] )
      THEN
        lrlMessErgebnis := rpMessErgebnis := 0;
        bpMessungOk := FALSE;
        blHelfer_RestwegMesung_Objekt_Gefunden := TRUE;
        lrlRestwegMessungMesstasterGefunden := l_mc_ReadActualPosition.Position;
      END_IF

    END_IF

  END_IF

END_IF
END_ACTION

(* ---- FreigabeEntziehen_Wiederanlauf.act.st ---- *)
(* METADATA
{
	"v3Meta": {
		"objectGuid": "91260ed7-d0f3-4853-b1f2-4ccb222d9ae8"
	}
}
*)
ACTION FreigabeEntziehen_Wiederanlauf
IF ( NOT blFreigabeEntziehenAktiv ) AND blFreigabeEntziehenAktivVorzyklus THEN
  // Reset-Freigabe erst nach aktivem Stop aufheben, sonst koennte rtlStop die Schrittkette unerwuenscht resetten.
  IF NOT blAchseStoppen AND NOT blAchseStoppenAktiv THEN
    blStopOhneReset := FALSE;
  END_IF

  // Wiederanlauf nach Pause:
  // Schritte ohne erneutes Execute := TRUE auf den jeweiligen Startschritt zuruecksetzen.
  CASE wlAktiveBetriebsart OF
    HANDPLUS:
      IF ( asteplSchritt[HANDPLUS] = STEP_400_E ) OR ( asteplSchritt[HANDPLUS] = STEP_1000_E ) THEN
        asteplSchritt[HANDPLUS] := STEP_300_E;
      END_IF

    HANDMINUS:
      IF ( asteplSchritt[HANDMINUS] = STEP_400_E ) OR ( asteplSchritt[HANDMINUS] = STEP_1000_E ) THEN
        asteplSchritt[HANDMINUS] := STEP_300_E;
      END_IF

    ABSOLUT:
      IF asteplSchritt[ABSOLUT] = STEP_500_E THEN
        asteplSchritt[ABSOLUT] := STEP_450_E;
      END_IF

    RELATIV:
      IF asteplSchritt[RELATIV] = STEP_500_E THEN
        asteplSchritt[RELATIV] := STEP_400_E;
      END_IF

    SCHEIBENMESSUNG:
      IF ( asteplSchritt[SCHEIBENMESSUNG] = STEP_350_E ) OR ( asteplSchritt[SCHEIBENMESSUNG] = STEP_500_E ) THEN
        asteplSchritt[SCHEIBENMESSUNG] := STEP_325_E;
      END_IF

    RESTWEG:
      IF asteplSchritt[RESTWEG] = STEP_450_E THEN
        asteplSchritt[RESTWEG] := STEP_400_E;
      ELSIF asteplSchritt[RESTWEG] = STEP_550_E THEN
        asteplSchritt[RESTWEG] := STEP_525_E;
      END_IF

    SYNC_AUF_MASTER:
      IF asteplSchritt[SYNC_AUF_MASTER] = STEP_1000_E THEN
        asteplSchritt[SYNC_AUF_MASTER] := STEP_400_E;
      END_IF

    INVERTIERTER_SYNC_AUF_MASTER:
      IF asteplSchritt[INVERTIERTER_SYNC_AUF_MASTER] = STEP_1000_E THEN
        asteplSchritt[INVERTIERTER_SYNC_AUF_MASTER] := STEP_400_E;
      END_IF

    RESET:
      IF asteplSchritt[RESET] = STEP_250_E THEN
        asteplSchritt[RESET] := STEP_200_E;
      ELSIF ( asteplSchritt[RESET] = STEP_325_E ) OR ( asteplSchritt[RESET] = STEP_350_E ) OR ( asteplSchritt[RESET] = STEP_400_E ) THEN
        asteplSchritt[RESET] := STEP_300_E;
      ELSIF ( asteplSchritt[RESET] = STEP_475_E ) OR ( asteplSchritt[RESET] = STEP_500_E ) THEN
        asteplSchritt[RESET] := STEP_450_E;
      END_IF
  END_CASE
END_IF

IF blFreigabeEntziehenAktiv THEN
  blStopOhneReset := TRUE;
  bpDone := FALSE;

  // Aktive MC-/CoE-Aktionen auch bei pausierter Betriebsartlogik sicher beenden
  l_fb_CoeLesen( i_b_Execute := FALSE );
  l_fb_CoeSchreiben( i_b_Execute := FALSE );
  l_mc_GearIn( Master := ppAntriebsInformationen.wAchsID, Slave := ppAntriebsInformationen.wAchsID, Execute := FALSE );
  l_mc_Reset( Axis := ppAntriebsInformationen.wAchsID, Execute := FALSE );
  l_mc_Home( Axis := ppAntriebsInformationen.wAchsID, Execute := FALSE );
  l_mc_MoveVelocity( Axis := ppAntriebsInformationen.wAchsID, Execute := FALSE );
  l_mc_MoveAbsolute( Axis := ppAntriebsInformationen.wAchsID, Execute := FALSE );

  // Warte-/Fehlertimer der eingefrorenen Schrittkette zuruecksetzen, damit die Haltezeit nicht als Timeout zaehlt
  tonlSoftwareFreigabe( IN := FALSE );
  tonlHardwareFreigabe( IN := FALSE );

  // Fahrtest nicht nur ueber bpAntrieblaeuft (Weg/Zyklus > 0.1 mm, 100 ms Entprellung -> langsame Fahrt / Anlauf wird als Stillstand gewertet),
  // sondern zusaetzlich ueber den MC-Status: Achse nicht im Stillstand (aber nicht Disabled/ungueltig) => MC_Stop, Power erst danach weg
  IF ( bpAntrieblaeuft OR bpAchseSychron OR l_mc_ReadStatus.Stopping OR blAchseStoppenAktiv
       OR ( l_mc_ReadStatus.Valid AND NOT l_mc_ReadStatus.StandStill AND NOT l_mc_ReadStatus.Disabled ) )
     AND NOT l_mc_ReadStatus.ErrorStop THEN
    blAchseStoppen := TRUE;
    blFreigabeEntziehenPowerAus := FALSE;
  ELSE
    blAchseStoppen := FALSE;
    blFreigabeEntziehenPowerAus := TRUE;
  END_IF
ELSE
  blFreigabeEntziehenPowerAus := FALSE;
END_IF
END_ACTION

(* ---- FUNKTION_Absolut_setzen.act.st ---- *)
(* METADATA
{
	"v3Meta": {
		"objectGuid": "5621efb7-cd40-4c15-9d03-482a92cbc1a2"
	}
}
*)
ACTION FUNKTION_Absolut_setzen
IF bpAbsolutSetzen THEN

  CASE asteplSchritt[ABSOLUT_SETZEN] OF

    STEP_0_E:
      bpAbsolutSetzenDone := FALSE;
      blReferenzLoeschen := TRUE; // Referenz ablöschen
      IF NOT bpIstReferenziert THEN
        blReferenzLoeschen := FALSE; // Referenz ablöschen
        asteplSchritt[ABSOLUT_SETZEN] := STEP_10_E;
      END_IF

    STEP_10_E:
      blReferenzSetzen := TRUE; //Referenz setzen
      IF bpIstReferenziert THEN
        blReferenzSetzen := FALSE;
        asteplSchritt[ABSOLUT_SETZEN] := STEP_1000_E;
      END_IF

    STEP_900_E:
      ;

    STEP_1000_E:
      bpAbsolutSetzenDone := TRUE;

  END_CASE

ELSE
  bpAbsolutSetzenDone := FALSE;
  blReferenzLoeschen := FALSE;
  blReferenzSetzen   := FALSE;
  asteplSchritt[ABSOLUT_SETZEN] := STEP_0_E;

END_IF
END_ACTION

(* ---- FUNKTION_Bremse_loesen.act.st ---- *)
(* METADATA
{
	"v3Meta": {
		"objectGuid": "8f122493-5427-4f74-8e27-0cfcccf91770"
	}
}
*)
ACTION FUNKTION_Bremse_loesen
IF bpBremseLoesen THEN

  CASE asteplSchritt[BREMSE_LOESEN] OF

    STEP_0_E:

      IF ppAntriebsInformationen.stOptionen.bBremseLoesenFreigabe THEN
        blBremseLoesen := TRUE; // Bremse lösen
        IF bpBremseGeloest THEN
          asteplSchritt[BREMSE_LOESEN] := STEP_1000_E;
        END_IF
      ELSE
        asteplSchritt[BREMSE_LOESEN] := STEP_900_E;
        blInternerFehler := TRUE;
        Antriebsfehler.wlBausteinFehlerNr := cKeineFreigabeZumBremseLoesen;
      END_IF

    STEP_900_E:
      ;

    STEP_1000_E:
      ;

  END_CASE

ELSE

  blBremseLoesen := FALSE;
  asteplSchritt[BREMSE_LOESEN] := STEP_0_E;

END_IF
END_ACTION

(* ---- Pruefe_Inputs_Langsamfahrt.act.st ---- *)
(* METADATA
{
	"v3Meta": {
		"objectGuid": "1b136394-d10a-4169-9faf-2f70a4dfcb82"
	}
}
*)
ACTION Pruefe_Inputs_Langsamfahrt
IF blZweiterZyklus OR blErsterZyklus THEN
  RETURN;
END_IF

rlGeschwindigkeit := rpGeschwindigkeit;
rlBeschleunigung  := rpBeschleunigung;
rlVerzoegerung    := rpVerzoegerung;

// Übergebene Geschwindigkeit über konfiguriertem Maximum
IF ( ( rlGeschwindigkeit ) > l_ts_MKAxisConfig.rVelocity / cFAKTOR_GESCHWINDIGKEIT_ECONSET ) THEN // EConSet in m/min angegeben...
  rlGeschwindigkeit := l_ts_MKAxisConfig.rVelocity / cFAKTOR_GESCHWINDIGKEIT_ECONSET;
END_IF
// Übergebene Geschwindigkeit kleiner 0
IF ( ( rlGeschwindigkeit ) < 0 ) THEN
  rlGeschwindigkeit := 0;
END_IF

// Übergebene Beschleunigung über konfiguriertem Maximum
IF ( ( rlBeschleunigung * cFAKTOR_RAMPEN ) > l_ts_MKAxisConfig.rAcceleration ) THEN
  rlBeschleunigung := l_ts_MKAxisConfig.rAcceleration / cFAKTOR_RAMPEN;
END_IF
// Übergebene Beschleunigung kleiner gleich 0
IF ( ( rlBeschleunigung * cFAKTOR_RAMPEN ) <= 0 ) THEN
  rlBeschleunigung := l_ts_MKAxisConfig.rAcceleration / cFAKTOR_RAMPEN;
END_IF

// Übergebene Verzögerung über konfiguriertem Maximum
IF ( ( rlVerzoegerung * cFAKTOR_RAMPEN ) > l_ts_MKAxisConfig.rDeceleration ) THEN
  rlVerzoegerung := l_ts_MKAxisConfig.rDeceleration / cFAKTOR_RAMPEN;
END_IF
// Übergebene Verzögerung kleiner gleich 0
IF ( ( rlVerzoegerung * cFAKTOR_RAMPEN ) <= 0 ) THEN
  rlVerzoegerung := l_ts_MKAxisConfig.rDeceleration / cFAKTOR_RAMPEN;
END_IF

// Wirksame Ruckzeit [s]: Vorgabe in ms, begrenzt durch EConSet.
rlRuckzeitSek := rpRuckzeit * 0.001;
IF rlRuckzeitSek <= 0 THEN
  rlRuckzeitSek := MAX(0.0, l_ts_MKAxisConfig.rRampTime);
ELSIF l_ts_MKAxisConfig.rRampTime > 0 THEN
  rlRuckzeitSek := MIN(rlRuckzeitSek, l_ts_MKAxisConfig.rRampTime);
END_IF

// Beide Jerk-Werte in MC-Einheiten bereitstellen.
// Welcher kleiner ist, haengt von Beschleunigung und Verzoegerung ab.
rlRuckBeschleunigung := 0;
rlRuckVerzoegerung := 0;
IF rlRuckzeitSek > 0 THEN
  rlRuckBeschleunigung := rlBeschleunigung * cFAKTOR_RAMPEN / rlRuckzeitSek;
  rlRuckVerzoegerung := rlVerzoegerung * cFAKTOR_RAMPEN / rlRuckzeitSek;
END_IF

// Die aktive Betriebsart waehlt danach in RuckFuerBewegung ihren Fahr-Jerk.
rlRuckzeit := rlRuckVerzoegerung;

/////////////////////////////////////////////////////////////////////////////////////////
/////////////////////////////////////////////////////////////////////////////////////////
// SHUTTLE LANGSAMFAHRT NOCKE
/////////////////////////////////////////////////////////////////////////////////////////
/////////////////////////////////////////////////////////////////////////////////////////
// Nocke in der aktuellen Fahrtrichtung erkennen.
blNockeInFahrtrichtung :=
                         (NOT udipEingaengeUmrichter.cXG31_2_I_2
                           AND eBewegungsrichtung = TE_Move_Direction.MD_NEGATIV_E)
                         OR (NOT udipEingaengeUmrichter.cXG31_1_I_1
                              AND eBewegungsrichtung = TE_Move_Direction.MD_POSITIV_E);

blEineLangsamfahrtnockeBelegt :=
                                NOT udipEingaengeUmrichter.cXG31_1_I_1
                                OR NOT udipEingaengeUmrichter.cXG31_2_I_2;

IF NOT bpAktiviereLangsamfahrtNocke
   OR rlGeschwindigkeit <=
   (l_ts_MKAxisConfig.rVelocity / cFAKTOR_GESCHWINDIGKEIT_ECONSET) * 0.1
THEN
  bpLangsamfahrenAktiv := FALSE;

ELSIF bpLangsamfahrenAktiv THEN
  // Bei kurz erkanntem Stillstand aktiv bleiben, solange eine Nocke belegt ist.
  bpLangsamfahrenAktiv :=
                         blNockeInFahrtrichtung
                         OR (eBewegungsrichtung = TE_Move_Direction.MD_STANDSTILL_E
                              AND blEineLangsamfahrtnockeBelegt);

ELSE
  // Während einer laufenden Verzögerung keine neue Langsamfahrt starten.
  bpLangsamfahrenAktiv :=
                         blNockeInFahrtrichtung AND NOT l_mc_ReadStatus.Decelerating;
END_IF
END_ACTION
